FOR u := 1 TO GVL_PARAM.UNIT_COUNT DO
	_stOut.astUnit[u].bPSetActive := FALSE;
END_FOR
IF i_nUnit >= 1 AND i_nUnit <= GVL_PARAM.UNIT_COUNT THEN
	_stOut.astUnit[i_nUnit].bPSetActive	:= i_bUnitPSetActive;
	_stOut.astUnit[i_nUnit].fPSet		:= i_fUnitPSet;
END_IF
// 새 지령: 값이 바뀌었거나 i_bSend
// [결함 13 수정 2026-11-04: 값 비교를 비트로 (운전원이 NaN을 넣어도 여기서 멈추지 않고 고르기에서 이상값으로 거름). 원래 _stOut.fPSet <> stOld.fPSet, _stOut.fQSet <> stOld.fQSet, …fPSet <> stOld.astUnit[u].fPSet]
_stOut.bNewSet := i_bSend
	OR _stOut.bPSetActive <> stOld.bPSetActive OR F_RealChanged(_stOut.fPSet, stOld.fPSet)
	OR _stOut.bQSetActive <> stOld.bQSetActive OR F_RealChanged(_stOut.fQSet, stOld.fQSet);
FOR u := 1 TO GVL_PARAM.UNIT_COUNT DO
	_stOut.bNewSet := _stOut.bNewSet
		OR _stOut.astUnit[u].bPSetActive <> stOld.astUnit[u].bPSetActive
		OR F_RealChanged(_stOut.astUnit[u].fPSet, stOld.astUnit[u].fPSet);
END_FOR
i_bSend := FALSE;

M_UpdateOutput := TRUE;		// 시험용: 항상 살아 있음 (만료 없음)
END_METHOD

END_FUNCTION_BLOCK

// ---- 20_Module/ControlMode/FB_CmPeakCut.TcPOU
FUNCTION_BLOCK FB_CmPeakCut EXTENDS FB_CmTariffBase		// 제어 모드: 피크컷 (Messis PEAK_SHAVING_MODE). 15분 평균 수전이 목표를 넘지 않게 방전
// 우선순위: 자동 충전 시간 → 잔량 방전 시간 (잔량 방전과 피크 제어 중 큰 값, 방전 허용 시간에만) → 피크 제어 (방전 허용 시간에만). 휴일·시각 무효 → 0
// 방전은 모두 역송 방지 (공통 설정). 피크 제어량 계산은 FB_CmPeakCalc (통합 모드와 같음)
VAR_INPUT
	i_stSet		: ST_CmPeakCutSet;		// 설정 (A_PassModuleSet이 GVL_PERSIST.g_stModuleSet.stCmPeakCut을 매 스캔 넘김)
END_VAR
VAR_OUTPUT
	q_fPeakCtrl	: REAL;		// 진단: 피크 제어량 (kW, FB_CmPeakCalc)
	q_nRemainMin	: UINT;		// 진단: 15분 구간 남은 분
	q_fExceeded	: REAL;		// 진단: 구간 목표 초과 수전 누적 (kW·분)
	q_fLoad1m	: REAL;		// 진단: 직전 1분 평균 부하 (kW)
END_VAR
VAR
	_fbPeak		: FB_CmPeakCalc;
END_VAR

METHOD M_Enter
VAR_INPUT
	i_stView	: ST_CtrlModeView;
END_VAR
SUPER^.M_Enter(i_stView := i_stView);
_fbPeak.M_Reset();
END_METHOD

METHOD M_Calc : ST_CtrlModeOut
VAR_INPUT
	i_stView	: ST_CtrlModeView;
END_VAR
VAR
	nNow	: UINT;
	fP		: REAL;
	fRem	: REAL;
	nRsn	: UINT;
	bNoCap	: BOOL;
END_VAR
fP := 0.0;
_fbPeak(i_stSet := i_stSet.stPeak, i_fRevMargin := i_stCommon.stNoRev.fMargin, i_stView := i_stView);		// 휴일에도 평균은 셈
q_fPeakCtrl		:= _fbPeak.q_fCtrl;
q_nRemainMin	:= _fbPeak.q_nRemainMin;
q_fExceeded		:= _fbPeak.q_fExceeded;
q_fLoad1m		:= _fbPeak.q_fLoad1m;
IF M_Begin(i_stView := i_stView) THEN
	nNow := F_TimeHhmm(i_stTime := i_stView.stTime);
	IF i_stSet.stAutoChg.bUse AND F_InHhmmWindow(i_nNow := nNow, i_nStart := i_stSet.stAutoChg.nStart, i_nEnd := i_stSet.stAutoChg.nEnd) THEN
		// 1) 자동 충전 (Messis MT_auto_charge)
		fP			:= -M_AutoChg(i_stView := i_stView, i_stWin := i_stSet.stAutoChg, q_bNoCap => bNoCap);
		q_nState	:= SEL(bNoCap, GVL_CM_RSN.AUTO_CHG, GVL_CM_RSN.NO_CAP);
	ELSIF i_stSet.stRemain.bUse AND F_InHhmmWindow(i_nNow := nNow, i_nStart := i_stSet.stRemain.nStart, i_nEnd := i_stSet.stRemain.nEnd) THEN
		// 2) 잔량 방전 (Messis MT_remain_discharge): 잔량 방전량이 있을 때만, 피크 제어량이 더 크면 그 값
		// [14번 수정 2026-11-09: 방전 허용 시간(공통 stDis: 시간·일요일) 밖이면 잔량 방전·피크 제어 모두 0, 상태 DIS_TIME.
		//   원래는 잔량 방전 시간이면 방전 허용 시간을 보지 않고 방전함]
		IF NOT M_DisAllowed(i_stTime := i_stView.stTime) THEN
			q_nState := GVL_CM_RSN.DIS_TIME;
		ELSE
			fRem		:= M_RemainDis(i_stView := i_stView, i_stWin := i_stSet.stRemain, q_bNoCap => bNoCap);
			q_nState	:= SEL(bNoCap, GVL_CM_RSN.REMAIN_DIS, GVL_CM_RSN.NO_CAP);
			IF fRem > 0.0 THEN
				fP := M_NoReverse(i_fReq := MAX(fRem, _fbPeak.q_fCtrl), i_stView := i_stView, q_nRsn => nRsn);
				IF nRsn <> 0 THEN
					q_nState := nRsn;
				END_IF
			END_IF
		END_IF
	ELSIF _fbPeak.q_bNewInterval THEN
		q_nState := GVL_CM_RSN.NEW_INTERVAL;
	ELSIF _fbPeak.q_fCtrl <= 0.0 THEN
		q_nState := GVL_CM_RSN.BELOW_PEAK;
	ELSIF NOT M_DisAllowed(i_stTime := i_stView.stTime) THEN
		q_nState := GVL_CM_RSN.DIS_TIME;
	ELSE
		// 3) 피크 제어 (Messis MT_peak_shaving_mode)
		fP			:= M_NoReverse(i_fReq := _fbPeak.q_fCtrl, i_stView := i_stView, q_nRsn => nRsn);
		q_nState	:= SEL(nRsn <> 0, GVL_CM_RSN.PEAK, nRsn);
	END_IF
END_IF
M_Calc := M_Finish(i_fP := fP);
END_METHOD

METHOD M_CheckSet : WSTRING(63)
M_CheckSet := SUPER^.M_CheckSet();
IF M_CheckSet <> "" THEN
	RETURN;
END_IF
// [결함 13 수정 2026-11-04: 피크 설정이 숫자인지 먼저]
IF NOT (F_RealOk(i_stSet.stPeak.fTarget) AND F_RealOk(i_stSet.stPeak.fBandSens) AND F_RealOk(i_stSet.stPeak.fLoadRatio) AND F_RealOk(i_stSet.stPeak.fMinOut)) THEN
	M_CheckSet := "피크컷: 피크 설정 숫자 아님";
ELSIF i_stSet.stPeak.fTarget < 0.0 OR i_stSet.stPeak.fBandSens < 0.0 OR i_stSet.stPeak.fLoadRatio < 0.0 OR i_stSet.stPeak.fLoadRatio > 1.0 OR i_stSet.stPeak.fMinOut < 0.0 THEN
	M_CheckSet := "피크컷: 목표·감도·부하 비율(0~1)·최소 출력";
ELSIF NOT M_CheckWindow(i_stWin := i_stSet.stAutoChg) THEN
	M_CheckSet := "피크컷: 자동 충전 시간·SOC";
ELSIF NOT M_CheckWindow(i_stWin := i_stSet.stRemain) THEN
	M_CheckSet := "피크컷: 잔량 방전 시간·SOC";
END_IF
END_METHOD

END_FUNCTION_BLOCK

// ---- 20_Module/ControlMode/FB_CmPeakCalc.TcPOU
FUNCTION_BLOCK FB_CmPeakCalc		// 15분 피크 제어량 계산 (Messis ACT_calc_quarter_avg_and_output 이식). 피크컷·통합 모드가 같이 씀
// 구간 = 시계 기준 15분 (매시 00·15·30·45분). 1초마다 수전·부하 평균, 시계 분이 바뀔 때마다 제어량 갱신, 구간 경계에서 0:
//   목표를 넘은 수전 누적 / 남은 분 (10 단위 반올림) × 속도 × (지난 분/15), 가용 출력 · 30초 평균 부하 × fLoadRatio · (30초 평균 부하 − 역송 여유) 상한
// 켜진 모드에서 매 스캔 부름. 모드가 켜질 때 M_Reset
VAR_INPUT
	i_stSet			: ST_CmPeakCalcSet;
	i_fRevMargin	: REAL;				// kW, 역송 방지 여유 (공통 설정 stNoRev.fMargin)
	i_stView		: ST_CtrlModeView;
END_VAR
VAR_OUTPUT
	q_fCtrl			: REAL;		// kW, 피크 제어 방전량 (0 = 제어 안 함). 1분마다 바뀜
	q_bNewInterval	: BOOL;		// 이번 스캔에 새 15분 구간 시작 (1스캔)
	q_nRemainMin	: UINT;		// 구간 남은 분
	q_fExceeded		: REAL;		// 이 구간 목표를 넘은 수전 누적 (kW·분)
	q_fLoad1m		: REAL;		// 직전 1분 평균 부하 (kW, ESS가 없을 때의 수전)
	q_bNoPcc		: BOOL;		// 접속점 계측 무효 (제어량 0, 평균 안 셈)
END_VAR
VAR
	_bInit			: BOOL;
	_nQuarter		: UINT;		// 지금 구간 번호 (시 × 4 + 분 / 15)
	_nPrevSec		: UINT;		// 지난 스캔 시계 초
	_nPrevMin		: UINT;		// 지난 스캔 시계 분
	_nPrevHalf		: UINT;		// 지난 스캔 30초 칸 (0 / 1)
	_n60			: UINT;		// 1분 평균 표본 수
	_n30			: UINT;		// 30초 평균 표본 수
	_fImp1m			: REAL;		// 1분 평균 수전 (kW)
	_fLoad30		: REAL;		// 30초 평균 부하 (kW)
	_fVelocity		: REAL;		// 제어 속도 (F_CmVelocity)
END_VAR
VAR_TEMP
	nQ				: UINT;
	fImp			: REAL;		// 수전 (kW)
	fLoad			: REAL;		// 부하 (kW)
	fCtrl			: REAL;
	nMin			: UINT;		// 구간 시작부터 지난 분
END_VAR

q_bNewInterval := FALSE;
q_bNoPcc := NOT i_stView.stGroup.stPcc.stMeas.stP.bValid;
IF NOT i_stView.stTime.bValid OR i_stSet.fTarget <= 0.0 THEN
	q_fCtrl	:= 0.0;
	_bInit	:= FALSE;
	RETURN;
END_IF

// 1) 구간 시작 (처음 또는 15분 경계). 경계에서는 제어량 0 (Messis: 남은 분 0으로 계산해 0)
nQ := i_stView.stTime.nHour * 4 + i_stView.stTime.nMinute / 15;
IF NOT _bInit OR nQ <> _nQuarter THEN
	q_bNewInterval	:= _bInit;		// 모드가 켜진 첫 스캔은 새 구간으로 보지 않음
	_bInit			:= TRUE;
	_nQuarter		:= nQ;
	_nPrevSec		:= i_stView.stTime.nSecond;
	_nPrevMin		:= i_stView.stTime.nMinute;
	_nPrevHalf		:= i_stView.stTime.nSecond / 30;
	_n60			:= 0;
	_n30			:= 0;
	q_nRemainMin	:= 15 - i_stView.stTime.nMinute MOD 15;
	q_fExceeded		:= 0.0;
	q_fCtrl			:= 0.0;
	_fVelocity		:= F_CmVelocity(i_fH := i_stSet.fTarget);
	RETURN;
END_IF

// 2) 시계의 초가 바뀔 때마다 (분·30초 경계는 시계 값으로 판단: 시계 보정으로 초가 건너뛰어도 밀리지 않음)
IF i_stView.stTime.nSecond <> _nPrevSec THEN
	_nPrevSec := i_stView.stTime.nSecond;
	// 3) 분이 바뀌면 지난 1분 평균으로 제어량 갱신
	IF i_stView.stTime.nMinute <> _nPrevMin THEN
		_nPrevMin		:= i_stView.stTime.nMinute;
		nMin			:= i_stView.stTime.nMinute MOD 15;		// 구간 시작부터 지난 분
		q_nRemainMin	:= 15 - nMin;
		fCtrl			:= 0.0;
		IF _n60 > 0 AND NOT q_bNoPcc THEN
			q_fExceeded := q_fExceeded + (_fImp1m - i_stSet.fTarget);
			IF q_fLoad1m - i_stSet.fTarget > i_stView.stGroup.fPRatedAvail * UINT_TO_REAL(q_nRemainMin / 15) * i_stSet.fBandSens * 0.5 THEN
				fCtrl := MIN(F_CmRoundTens(i_f := q_fExceeded / UINT_TO_REAL(q_nRemainMin)) * _fVelocity * (UINT_TO_REAL(nMin) / 15.0), i_stView.stGroup.fPRatedAvail);
			END_IF
			fCtrl := MIN(fCtrl, _fLoad30 * i_stSet.fLoadRatio);
			fCtrl := MIN(fCtrl, _fLoad30 - i_fRevMargin);
			IF fCtrl <= 1.0 THEN
				fCtrl := 0.0;
			ELSE
				fCtrl := MAX(fCtrl, i_stSet.fMinOut);
			END_IF
			IF _fImp1m - i_stSet.fTarget > 0.0 THEN
				_fVelocity := F_CmVelocity(i_fH := _fImp1m - i_stSet.fTarget);
			END_IF
		END_IF
		q_fCtrl	:= fCtrl;
		_n60	:= 0;			// 다음 1분 평균을 새로 셈 (값은 남김)
	END_IF
	IF i_stView.stTime.nSecond / 30 <> _nPrevHalf THEN
		_nPrevHalf	:= i_stView.stTime.nSecond / 30;
		_n30		:= 0;		// 다음 30초 평균을 새로 셈 (값은 남김)
	END_IF
	// 4) 1초 표본
	IF q_bNoPcc THEN
		q_fCtrl := 0.0;			// 계측 무효: 평균에 넣지 않고 제어 안 함
	ELSE
		_n60	:= _n60 + 1;
		_n30	:= _n30 + 1;
		fImp	:= -i_stView.stGroup.stPcc.stMeas.stP.fValue;			// 수전 + (접속점 P는 공급 +)
		fLoad	:= i_stView.stGroup.fPOut + fImp;							// ESS가 없을 때의 수전
		_fImp1m		:= (_fImp1m * UINT_TO_REAL(_n60 - 1) + fImp) / UINT_TO_REAL(_n60);
		q_fLoad1m	:= (q_fLoad1m * UINT_TO_REAL(_n60 - 1) + fLoad) / UINT_TO_REAL(_n60);
		_fLoad30	:= (_fLoad30 * UINT_TO_REAL(_n30 - 1) + fLoad) / UINT_TO_REAL(_n30);
	END_IF
END_IF

METHOD M_Reset		// 모드가 켜질 때: 구간을 지금부터 다시 셈, 제어량 0
_bInit		:= FALSE;
q_fCtrl		:= 0.0;
q_fExceeded	:= 0.0;
q_fLoad1m	:= 0.0;
_fImp1m		:= 0.0;
_fLoad30	:= 0.0;
END_METHOD

END_FUNCTION_BLOCK

// ---- 20_Module/ControlMode/F_CmVelocity.TcPOU
FUNCTION F_CmVelocity : REAL		// 피크 제어 속도 (Messis getVelocity): 넘는 양이 작을수록 크게. (log10(h + 100) − log10(h)) × 20, h ≤ 0이면 1
VAR_INPUT
	i_fH		: REAL;		// kW, 목표 또는 목표를 넘은 양
END_VAR

IF i_fH <= 0.0 THEN
	F_CmVelocity := 1.0;
ELSE
	F_CmVelocity := (LOG(i_fH + 100.0) - LOG(i_fH)) * 20.0;
END_IF

END_FUNCTION

// ---- 20_Module/ControlMode/F_CmRoundTens.TcPOU
FUNCTION F_CmRoundTens : REAL		// 10 단위 반올림 (Messis roundUpTens)
VAR_INPUT
	i_f			: REAL;
END_VAR

// [결함 13 수정 2026-11-04: NaN·범위 밖이면 REAL_TO_DINT가 FPU 예외 → F_RealToDint (NaN은 0). 원래 DINT_TO_REAL(REAL_TO_DINT(i_f / 10.0)) * 10.0]
F_CmRoundTens := DINT_TO_REAL(F_RealToDint(i_f / 10.0)) * 10.0;

END_FUNCTION

// ---- 20_Module/ControlMode/FB_CmSchedPeak.TcPOU
FUNCTION_BLOCK FB_CmSchedPeak EXTENDS FB_CmTariffBase		// 제어 모드: 통합 = 스케줄 + 피크컷 (Messis SCHEDULE_PS_MODE)
// 우선순위: 잔량 방전 시간 (잔량 방전과 피크 제어 중 큰 값, 방전 허용 시간에만) → 피크 제어가 필요하고 방전 허용 시간이면 (피크 제어량과 시간표 방전 중 큰 값)
//   → 아니면 스케줄 모드와 같음. 시간표는 스케줄 모드와 같은 표, 피크 제어량 계산은 피크컷과 같은 FB_CmPeakCalc
// Messis와 다른 점: 시간표가 충전 칸일 때 피크 제어가 필요하면 피크 제어량만 방전 (Messis는 충전값 크기만큼 방전할 수 있었음)
VAR_INPUT
	i_stTable	: ST_CmScheduleSet;		// 시간표 (스케줄 모드와 같은 GVL_PERSIST.g_stModuleSet.stCmSchedule)
	i_stSet		: ST_CmSchedPeakSet;	// 설정 (GVL_PERSIST.g_stModuleSet.stCmSchedPeak)
END_VAR
VAR_OUTPUT
	q_fPeakCtrl	: REAL;		// 진단: 피크 제어량 (kW, FB_CmPeakCalc)
	q_nRemainMin	: UINT;		// 진단: 15분 구간 남은 분
	q_fExceeded	: REAL;		// 진단: 구간 목표 초과 수전 누적 (kW·분)
	q_fLoad1m	: REAL;		// 진단: 직전 1분 평균 부하 (kW)
END_VAR
VAR
	_fbPeak		: FB_CmPeakCalc;
END_VAR

METHOD M_Enter
VAR_INPUT
	i_stView	: ST_CtrlModeView;
END_VAR
SUPER^.M_Enter(i_stView := i_stView);
_fbPeak.M_Reset();
END_METHOD

METHOD M_Calc : ST_CtrlModeOut
VAR_INPUT
	i_stView	: ST_CtrlModeView;
END_VAR
VAR
	nNow	: UINT;
	fP		: REAL;
	fRem	: REAL;
	nRsn	: UINT;
	bNoCap	: BOOL;
END_VAR
fP := 0.0;
_fbPeak(i_stSet := i_stSet.stPeak, i_fRevMargin := i_stCommon.stNoRev.fMargin, i_stView := i_stView);
q_fPeakCtrl		:= _fbPeak.q_fCtrl;
q_nRemainMin	:= _fbPeak.q_nRemainMin;
q_fExceeded		:= _fbPeak.q_fExceeded;
q_fLoad1m		:= _fbPeak.q_fLoad1m;
IF M_Begin(i_stView := i_stView) THEN
	nNow := F_TimeHhmm(i_stTime := i_stView.stTime);
	M_SchedLookup(i_stTime := i_stView.stTime, iq_stTable := i_stTable);
	IF i_stSet.stRemain.bUse AND F_InHhmmWindow(i_nNow := nNow, i_nStart := i_stSet.stRemain.nStart, i_nEnd := i_stSet.stRemain.nEnd) THEN
		// 1) 잔량 방전
		// [14번 수정 2026-11-09: 방전 허용 시간(공통 stDis: 시간·일요일) 밖이면 잔량 방전·피크 제어 모두 0, 상태 DIS_TIME.
		//   원래는 잔량 방전 시간이면 방전 허용 시간을 보지 않고 방전함]
		IF NOT M_DisAllowed(i_stTime := i_stView.stTime) THEN
			q_nState := GVL_CM_RSN.DIS_TIME;
		ELSE
			fRem		:= M_RemainDis(i_stView := i_stView, i_stWin := i_stSet.stRemain, q_bNoCap => bNoCap);
			q_nState	:= SEL(bNoCap, GVL_CM_RSN.REMAIN_DIS, GVL_CM_RSN.NO_CAP);
			IF fRem > 0.0 THEN
				fP := M_NoReverse(i_fReq := MAX(fRem, _fbPeak.q_fCtrl), i_stView := i_stView, q_nRsn => nRsn);
				IF nRsn <> 0 THEN
					q_nState := nRsn;
				END_IF
			END_IF
		END_IF
	ELSIF _fbPeak.q_fCtrl > 0.0 AND M_DisAllowed(i_stTime := i_stView.stTime) THEN
		// 2) 피크 제어 + 시간표 방전 중 큰 값
		fP			:= M_NoReverse(i_fReq := MAX(_fbPeak.q_fCtrl, MAX(q_fSlotP, 0.0)), i_stView := i_stView, q_nRsn => nRsn);
		q_nState	:= SEL(nRsn <> 0, GVL_CM_RSN.SCHED_PEAK, nRsn);
	ELSE
		// 3) 스케줄만
		fP			:= M_SchedOut(i_stView := i_stView, q_nRsn => nRsn);
		q_nState	:= nRsn;
	END_IF
END_IF
M_Calc := M_Finish(i_fP := fP);
END_METHOD

METHOD M_CheckSet : WSTRING(63)
M_CheckSet := SUPER^.M_CheckSet();
IF M_CheckSet <> "" THEN
	RETURN;
END_IF
M_CheckSet := M_CheckTable(iq_stTable := i_stTable);
IF M_CheckSet <> "" THEN
	RETURN;
END_IF
// [결함 13 수정 2026-11-04: 피크 설정이 숫자인지 먼저]
IF NOT (F_RealOk(i_stSet.stPeak.fTarget) AND F_RealOk(i_stSet.stPeak.fBandSens) AND F_RealOk(i_stSet.stPeak.fLoadRatio) AND F_RealOk(i_stSet.stPeak.fMinOut)) THEN
	M_CheckSet := "통합: 피크 설정 숫자 아님";
ELSIF i_stSet.stPeak.fTarget < 0.0 OR i_stSet.stPeak.fBandSens < 0.0 OR i_stSet.stPeak.fLoadRatio < 0.0 OR i_stSet.stPeak.fLoadRatio > 1.0 OR i_stSet.stPeak.fMinOut < 0.0 THEN
	M_CheckSet := "통합: 목표·감도·부하 비율(0~1)·최소 출력";
ELSIF NOT M_CheckWindow(i_stWin := i_stSet.stRemain) THEN
	M_CheckSet := "통합: 잔량 방전 시간·SOC";
END_IF
END_METHOD

END_FUNCTION_BLOCK

// ---- 20_Module/Common/FB_SocLimit.TcPOU
FUNCTION_BLOCK FB_SocLimit EXTENDS FB_ModuleBase IMPLEMENTS I_BatLimitRule	// SOC 감발·차단·재개 마진 (버스 제한). 기본 SOC 정책 (Auto·Manual 기본 등록)
// 최대 SOC가 상한에 다가가면 충전 한도를, 최소 SOC가 하한에 다가가면 방전 한도를 줄이고, 한계에서 막음
// 막은 뒤에는 SOC가 재개 마진만큼 돌아와야 다시 허용. 다시 허용한 뒤 감발 구간을 지나는 동안 bResume (재개 램프율)
// 출력 한도만 냄 (장비 명령 없음). 한도가 0이면 그 방향 출력 0 = 대기
// nTarget 0 = 모든 버스를 한 인스턴스가 봄 (버스마다 상태를 따로 가짐)
VAR_INPUT
	i_stSet	: ST_SocLimitSet;	// 설정 (MAIN이 GVL_PERSIST.g_stModuleSet 칸을 매 스캔 넘김. 안 넘기면 기본값)
END_VAR
VAR
	(* 버스마다 상태 *)
	_abChgBlock	: ARRAY[1..GVL_PARAM.BAT_COUNT] OF BOOL;	// 충전 막음 (재개 마진 전까지 유지)
	_abDisBlock	: ARRAY[1..GVL_PARAM.BAT_COUNT] OF BOOL;	// 방전 막음
	_abChgResume	: ARRAY[1..GVL_PARAM.BAT_COUNT] OF BOOL;	// 충전 재개 중 (막음이 풀린 뒤 감발 구간)
	_abDisResume	: ARRAY[1..GVL_PARAM.BAT_COUNT] OF BOOL;
	_afChgRatio	: ARRAY[1..GVL_PARAM.BAT_COUNT] OF REAL;	// 진단: 충전 한도 비율 (1 = 안 줄임)
	_afDisRatio	: ARRAY[1..GVL_PARAM.BAT_COUNT] OF REAL;	// 진단: 방전 한도 비율
END_VAR
VAR CONSTANT
	RSN_CHG_DERATE	: UINT := 1;	// 상한 근처 충전 감발
	RSN_CHG_BLOCK	: UINT := 2;	// 상한 충전 막음
	RSN_DIS_DERATE	: UINT := 3;	// 하한 근처 방전 감발
	RSN_DIS_BLOCK	: UINT := 4;	// 하한 방전 막음
	RSN_SOC_INVALID	: UINT := 5;	// SOC 무효
END_VAR

METHOD M_Evaluate : ST_BatLimitOut
VAR_INPUT
	i_stView	: ST_BatLimitView;
END_VAR
VAR
	b	: UINT;
	fChg	: REAL;	// 충전 한도 비율
	fDis	: REAL;	// 방전 한도 비율
END_VAR
b := i_stView.nBatGroup;
IF b < 1 OR b > GVL_PARAM.BAT_COUNT THEN
	RETURN;
END_IF
// SOC 무효: 상태를 풀고, 설정이면 충·방전 모두 막음
IF NOT i_stView.stSocMax.bValid OR NOT i_stView.stSocMin.bValid THEN
	_abChgBlock[b]	:= FALSE;
	_abDisBlock[b]	:= FALSE;
	_abChgResume[b]	:= FALSE;
	_abDisResume[b]	:= FALSE;
	_afChgRatio[b]	:= 1.0;
	_afDisRatio[b]	:= 1.0;
	IF i_stSet.bBlockOnInvalid THEN
		M_Evaluate.stP.bActive	:= TRUE;
		M_Evaluate.stP.fMax	:= 0.0;
		M_Evaluate.stP.fMin	:= 0.0;
		M_Evaluate.stP.nReason	:= RSN_SOC_INVALID;
		_afChgRatio[b]	:= 0.0;
		_afDisRatio[b]	:= 0.0;
	END_IF
	RETURN;
END_IF

// 충전: 최대 SOC 기준
IF i_stView.stSocMax.fValue >= i_stSet.fSocMax THEN
	_abChgBlock[b]	:= TRUE;
	_abChgResume[b]	:= FALSE;
ELSIF _abChgBlock[b] AND i_stView.stSocMax.fValue <= i_stSet.fSocMax - i_stSet.fResumeMargin THEN
	_abChgBlock[b]	:= FALSE;
	_abChgResume[b]	:= TRUE;
END_IF
fChg := 0.0;
IF NOT _abChgBlock[b] THEN
	fChg := F_SocDerate(i_fSoc := i_stView.stSocMax.fValue, i_fLimit := i_stSet.fSocMax, i_fBand := i_stSet.fBand, i_bUpper := TRUE);
END_IF
IF fChg >= 1.0 THEN
	_abChgResume[b] := FALSE;
END_IF

// 방전: 최소 SOC 기준
IF i_stView.stSocMin.fValue <= i_stSet.fSocMin THEN
	_abDisBlock[b]	:= TRUE;
	_abDisResume[b]	:= FALSE;
ELSIF _abDisBlock[b] AND i_stView.stSocMin.fValue >= i_stSet.fSocMin + i_stSet.fResumeMargin THEN
	_abDisBlock[b]	:= FALSE;
	_abDisResume[b]	:= TRUE;
END_IF
fDis := 0.0;
IF NOT _abDisBlock[b] THEN
	fDis := F_SocDerate(i_fSoc := i_stView.stSocMin.fValue, i_fLimit := i_stSet.fSocMin, i_fBand := i_stSet.fBand, i_bUpper := FALSE);
END_IF
IF fDis >= 1.0 THEN
	_abDisResume[b] := FALSE;
END_IF

_afChgRatio[b]	:= fChg;
_afDisRatio[b]	:= fDis;
M_Evaluate.bResume := _abChgResume[b] OR _abDisResume[b];
IF fChg < 1.0 OR fDis < 1.0 THEN
	M_Evaluate.stP.bActive	:= TRUE;
	M_Evaluate.stP.fMax	:= MAX(i_stView.fPDisMax, 0.0) * fDis;
	M_Evaluate.stP.fMin	:= -MAX(i_stView.fPChgMax, 0.0) * fChg;
	// 이유: 막음이 감발보다 먼저 (한 줄 제한이라 상·하한이 같은 이유를 가짐)
	IF _abDisBlock[b] THEN
		M_Evaluate.stP.nReason := RSN_DIS_BLOCK;
	ELSIF _abChgBlock[b] THEN
		M_Evaluate.stP.nReason := RSN_CHG_BLOCK;
	ELSIF fDis < 1.0 THEN
		M_Evaluate.stP.nReason := RSN_DIS_DERATE;
	ELSE
		M_Evaluate.stP.nReason := RSN_CHG_DERATE;
	END_IF
END_IF
END_METHOD

METHOD M_ReasonText : WSTRING(63)
VAR_INPUT
	i_nReason	: UINT;
END_VAR
CASE i_nReason OF
	RSN_CHG_DERATE:	M_ReasonText := "SOC 상한 근처 충전 감발";
	RSN_CHG_BLOCK:	M_ReasonText := "SOC 상한 충전 막음";
	RSN_DIS_DERATE:	M_ReasonText := "SOC 하한 근처 방전 감발";
	RSN_DIS_BLOCK:	M_ReasonText := "SOC 하한 방전 막음";
	RSN_SOC_INVALID:	M_ReasonText := "SOC 무효";
ELSE
	M_ReasonText := WCONCAT("이유 ", TO_WSTRING(i_nReason));
END_CASE
END_METHOD

METHOD M_CheckSet : WSTRING(63)		// 설정 점검: SOC 상·하한, 감발 폭, 재개 마진
// [9-21 수정 2026-11-04: 검사 규칙을 F_SocLimitSetErr로 옮김 (EMS config 반영 FB_EmsConfigApply와 같은 규칙을 씀). 원래:
//   M_CheckSet := "";
//   IF NOT (F_RealOk(i_stSet.fSocMin) AND F_RealOk(i_stSet.fSocMax) AND F_RealOk(i_stSet.fBand) AND F_RealOk(i_stSet.fResumeMargin)) THEN	// [결함 13 수정 2026-11-04]
//   	M_CheckSet := "SOC 설정 숫자 아님";
//   ELSIF i_stSet.fSocMin < 0.0 OR i_stSet.fSocMax > 100.0 OR i_stSet.fSocMin >= i_stSet.fSocMax THEN
//   	M_CheckSet := "SOC 상·하한 (0 ≤ 하한 < 상한 ≤ 100)";
//   ELSIF i_stSet.fBand < 0.0 OR i_stSet.fSocMin + i_stSet.fBand > i_stSet.fSocMax - i_stSet.fBand THEN
//   	M_CheckSet := "감발 폭 fBand (0 이상, 상·하한 사이)";
//   ELSIF i_stSet.fResumeMargin < 0.0 OR i_stSet.fSocMin + i_stSet.fResumeMargin >= i_stSet.fSocMax - i_stSet.fResumeMargin THEN
//   	M_CheckSet := "재개 마진 fResumeMargin (0 이상, 상·하한 사이)";
//   END_IF]
M_CheckSet := F_SocLimitSetErr(i_stSet);
END_METHOD

END_FUNCTION_BLOCK

// ---- 20_Module/Common/F_SocDerate.TcPOU
FUNCTION F_SocDerate : REAL	// SOC 감발 비율 (0~1, 상태 없음). 여러 SOC 정책 모듈이 같이 씀
// 상한(i_bUpper = TRUE, 충전 쪽): SOC ≥ 한계면 0, 한계 - 폭 < SOC면 선형으로 줄임, 그 아래는 1
// 하한(i_bUpper = FALSE, 방전 쪽): SOC ≤ 한계면 0, SOC < 한계 + 폭이면 선형으로 줄임, 그 위는 1
VAR_INPUT
	i_fSoc	: REAL;	// %
	i_fLimit	: REAL;	// %, 한계
	i_fBand	: REAL;	// %, 감발 폭. 0 이하면 줄이지 않고 한계에서 0
	i_bUpper	: BOOL;	// TRUE = 상한, FALSE = 하한
END_VAR

IF i_bUpper THEN
	IF i_fSoc >= i_fLimit THEN
		F_SocDerate := 0.0;
	ELSIF i_fBand > 0 AND i_fSoc > i_fLimit - i_fBand THEN
		F_SocDerate := (i_fLimit - i_fSoc) / i_fBand;
	ELSE
		F_SocDerate := 1.0;
	END_IF
ELSE
	IF i_fSoc <= i_fLimit THEN
		F_SocDerate := 0.0;
	ELSIF i_fBand > 0 AND i_fSoc < i_fLimit + i_fBand THEN
		F_SocDerate := (i_fSoc - i_fLimit) / i_fBand;
	ELSE
		F_SocDerate := 1.0;
	END_IF
END_IF

END_FUNCTION

// ---- 20_Module/Common/FB_UnitLimit.TcPOU
FUNCTION_BLOCK FB_UnitLimit EXTENDS FB_ModuleBase IMPLEMENTS I_UnitLimitRule	// 사용자 한도: 유닛마다 운전원이 정한 P·Q 상·하한 (kW·kvar). 정격·Derate와 겹쳐 좁은 쪽 (코어 FB_EquipmentLimits)
// 등록: g_aipUnitRule 한 칸, g_astUnitRuleReg nTarget 0 (전체 유닛, 유닛마다 설정을 따로 봄), bAuto·bManual로 적용 모드
// 출력 제한 이유: 유닛 한도 UnitRule + 이 모듈 ID, 이유 "사용자 한도"
VAR_INPUT
	i_stSet		: ST_UnitLimitSet;	// 유닛마다 한도 (MAIN A_PassModuleSet이 g_stModuleSet 칸을 넘김. 안 넘기면 모두 끔)
END_VAR
VAR CONSTANT
	RSN_USER	: UINT := 1;		// 사용자 한도
END_VAR

METHOD M_Evaluate : ST_LimitOut
VAR_INPUT
	i_stView	: ST_UnitLimitView;
END_VAR
VAR
	u	: UINT;
END_VAR
u := i_stView.nUnit;
IF u < 1 OR u > GVL_PARAM.UNIT_COUNT THEN
	RETURN;
END_IF
IF i_stSet.astUnit[u].bPEnable THEN
	M_Evaluate.stP.bActive	:= TRUE;
	M_Evaluate.stP.fMax		:= i_stSet.astUnit[u].fPMax;
	M_Evaluate.stP.fMin		:= i_stSet.astUnit[u].fPMin;
	M_Evaluate.stP.nReason	:= RSN_USER;
END_IF
IF i_stSet.astUnit[u].bQEnable THEN
	M_Evaluate.stQ.bActive	:= TRUE;
	M_Evaluate.stQ.fMax		:= i_stSet.astUnit[u].fQMax;
	M_Evaluate.stQ.fMin		:= i_stSet.astUnit[u].fQMin;
	M_Evaluate.stQ.nReason	:= RSN_USER;
END_IF
END_METHOD

METHOD M_ReasonText : WSTRING(63)
VAR_INPUT
	i_nReason	: UINT;
END_VAR
IF i_nReason = RSN_USER THEN
	M_ReasonText := "사용자 한도";
ELSE
	M_ReasonText := WCONCAT("이유 ", TO_WSTRING(i_nReason));
END_IF
END_METHOD

METHOD M_CheckSet : WSTRING(63)		// 설정 점검: 켠 한도는 상한 ≥ 0 ≥ 하한
VAR
	u	: UINT;
END_VAR
M_CheckSet := "";
FOR u := 1 TO GVL_PARAM.UNIT_COUNT DO
	IF NOT (F_RealOk(i_stSet.astUnit[u].fPMax) AND F_RealOk(i_stSet.astUnit[u].fPMin) AND F_RealOk(i_stSet.astUnit[u].fQMax) AND F_RealOk(i_stSet.astUnit[u].fQMin)) THEN	// [결함 13 수정 2026-11-04]
		M_CheckSet := F_TxtNum("한도 숫자 아님: 유닛 ", u);
		RETURN;
	END_IF
	IF i_stSet.astUnit[u].bPEnable AND (i_stSet.astUnit[u].fPMax < 0.0 OR i_stSet.astUnit[u].fPMin > 0.0) THEN
		M_CheckSet := F_TxtNum("P 한도 상한 < 0 또는 하한 > 0: 유닛 ", u);
		RETURN;
	END_IF
	IF i_stSet.astUnit[u].bQEnable AND (i_stSet.astUnit[u].fQMax < 0.0 OR i_stSet.astUnit[u].fQMin > 0.0) THEN
		M_CheckSet := F_TxtNum("Q 한도 상한 < 0 또는 하한 > 0: 유닛 ", u);
		RETURN;
	END_IF
END_FOR
END_METHOD

END_FUNCTION_BLOCK

// ---- 20_Module/Standard/FB_ProtPcsFault.TcPOU
FUNCTION_BLOCK FB_ProtPcsFault EXTENDS FB_ModuleBase IMPLEMENTS I_ProtectionRule		// 표준 보호: PCS 고장 (범위 Unit): 통신이 있고 PCS가 고장을 알림. 기본 등록. 빼면 이 보호 없음. 현장마다 다르면 복사해 이름을 바꿔 그 칸에 대신 등록
VAR
END_VAR

METHOD M_Evaluate : BOOL		// 범위가 맞지 않게 등록되면 FALSE (보호 안 걸림)
VAR_INPUT
	i_stView	: ST_ProtView;
END_VAR
M_Evaluate := i_stView.eScope = E_ProtScope.Unit AND i_stView.bInstalled AND i_stView.stUnit.bComm AND i_stView.stUnit.bFault;
END_METHOD

END_FUNCTION_BLOCK

// ---- 20_Module/Standard/FB_ProtPcsComm.TcPOU
FUNCTION_BLOCK FB_ProtPcsComm EXTENDS FB_ModuleBase IMPLEMENTS I_ProtectionRule		// 표준 보호: PCS 통신 끊김 (범위 Unit). 기본 등록. 빼면 이 보호 없음. 현장마다 다르면 복사해 이름을 바꿔 그 칸에 대신 등록
VAR
END_VAR

METHOD M_Evaluate : BOOL		// 범위가 맞지 않게 등록되면 FALSE (보호 안 걸림)
VAR_INPUT
	i_stView	: ST_ProtView;
END_VAR
M_Evaluate := i_stView.eScope = E_ProtScope.Unit AND i_stView.bInstalled AND NOT i_stView.stUnit.bComm;
END_METHOD

END_FUNCTION_BLOCK

// ---- 20_Module/Standard/FB_ProtBmsFault.TcPOU
FUNCTION_BLOCK FB_ProtBmsFault EXTENDS FB_ModuleBase IMPLEMENTS I_ProtectionRule		// 표준 보호: BMS 고장 (범위 Bms): 통신이 있고 BMS가 고장을 알림. 기본 등록. 빼면 이 보호 없음. 현장마다 다르면 복사해 이름을 바꿔 그 칸에 대신 등록
VAR
END_VAR

METHOD M_Evaluate : BOOL		// 범위가 맞지 않게 등록되면 FALSE (보호 안 걸림)
VAR_INPUT
	i_stView	: ST_ProtView;
END_VAR
M_Evaluate := i_stView.eScope = E_ProtScope.Bms AND i_stView.bInstalled AND i_stView.stBms.bComm AND i_stView.stBms.bFault;
END_METHOD

END_FUNCTION_BLOCK

// ---- 20_Module/Standard/FB_ProtBmsComm.TcPOU
FUNCTION_BLOCK FB_ProtBmsComm EXTENDS FB_ModuleBase IMPLEMENTS I_ProtectionRule		// 표준 보호: BMS 통신 끊김 (범위 Bms). 기본 등록. 빼면 이 보호 없음. 현장마다 다르면 복사해 이름을 바꿔 그 칸에 대신 등록
VAR
END_VAR

METHOD M_Evaluate : BOOL		// 범위가 맞지 않게 등록되면 FALSE (보호 안 걸림)
VAR_INPUT
	i_stView	: ST_ProtView;
END_VAR
M_Evaluate := i_stView.eScope = E_ProtScope.Bms AND i_stView.bInstalled AND NOT i_stView.stBms.bComm;
END_METHOD

END_FUNCTION_BLOCK

// ---- 20_Module/Standard/FB_ProtPccInvalid.TcPOU
FUNCTION_BLOCK FB_ProtPccInvalid EXTENDS FB_ModuleBase IMPLEMENTS I_ProtectionRule		// 표준 보호: 접속점 계측 무효 (범위 Group): 접속점 유효전력 값이 무효. 기본 등록. 빼면 이 보호 없음. 현장마다 다르면 복사해 이름을 바꿔 그 칸에 대신 등록
VAR
END_VAR

METHOD M_Evaluate : BOOL		// 범위가 맞지 않게 등록되면 FALSE (보호 안 걸림)
VAR_INPUT
	i_stView	: ST_ProtView;
END_VAR
// [결함 7 수정 2026-11-03: 접속점이 없는 그룹(nPccPoint 0)은 판단 안 함. 원래 M_Evaluate := i_stView.eScope = E_ProtScope.Group AND NOT i_stView.stPcc.stMeas.stP.bValid;]
M_Evaluate := i_stView.eScope = E_ProtScope.Group AND NOT i_stView.stPcc.bNoPoint AND NOT i_stView.stPcc.stMeas.stP.bValid;
END_METHOD

END_FUNCTION_BLOCK

// ---- 20_Module/Standard/FB_ProtRespStd.TcPOU
FUNCTION_BLOCK FB_ProtRespStd EXTENDS FB_ModuleBase IMPLEMENTS I_ProtResponse		// 표준 보호 대응 (기본 등록: GVL_SITE.g_aipResp 칸마다 같은 인스턴스): 칸 설정(ST_ProtCfg)의 조치를 범위 안 유닛·BMS에 한 단계로 요청
// 유닛: 범위에 드는 유닛 중 그 운전 모드에 조치를 거는 것(bAuto·bManual)만. 모드 조치(ToManual)는 bAuto 항목이면 범위 안 유닛 전부
// BMS: Bms·BatGroup 범위는 그 버스에 조치를 받는 유닛이 있을 때 (버스에 유닛이 없으면 그대로). Unit·Group·Site 범위는 조치를 받는 유닛의 배터리 그룹 BMS 전부
// 현장 대응이 다르면 이 FB를 복사해 이름을 바꿔 그 칸에 대신 등록. 상태가 없어 인스턴스 하나를 모든 칸에 같이 등록함

METHOD M_Respond		// 칸 설정(stProt)의 조치를 걸렸을 때만 요청
// 코어가 매 스캔 범위 안 대상마다 부름 (조건이 없을 때도: 단계 대응의 타이머·상태를 풀 수 있게). 대상 번호가 0으로 등록되면 대상마다 상태를 따로 둠
VAR_INPUT
	i_bActive		: BOOL;			// 보호 조건 있음 (등록 bAuto·bManual 중 하나가 켜져 있고 조건 모듈이 TRUE)
	i_tActive		: TIME;			// 조건이 이어진 시간 (조건 없으면 0)
	i_nTarget		: UINT;			// 대상 번호 (범위는 i_stRule.eScope. Site면 1)
	i_stRule		: ST_RuleCfg;		// 이 칸 설정 (범위·대상·임계값·표준 대응 설정)
END_VAR
VAR_IN_OUT CONSTANT
	iq_astUnit		: ARRAY[1..GVL_PARAM.UNIT_COUNT] OF ST_UnitState;	// 장비 상태 (이번 스캔 스냅샷, 읽기 전용)
	iq_astBms		: ARRAY[1..GVL_PARAM.BMS_COUNT] OF ST_BatState;
	iq_astUnitCfg	: ARRAY[1..GVL_PARAM.UNIT_COUNT] OF ST_UnitCfg;		// 소속 (제어 그룹·배터리 그룹)
	iq_astBmsCfg	: ARRAY[1..GVL_PARAM.BMS_COUNT] OF ST_BmsCfg;
	iq_aeOpMode		: ARRAY[1..GVL_PARAM.UNIT_COUNT] OF E_OpMode;		// 실제 운전 모드
END_VAR
VAR_IN_OUT
	iq_stReq		: ST_ProtReq;		// 요청 (코어가 비워서 넘김)
END_VAR
VAR
	u			: UINT;
	m			: UINT;
	nBus		: UINT;		// Bms·BatGroup 범위의 배터리 그룹
	nBusUnits	: UINT;		// 그 버스의 유닛 수
	bBusTakes	: BOOL;		// 그 버스에 조치를 받는 유닛이 있음
	bIn			: BOOL;
	bManual		: BOOL;
	bTakes		: BOOL;
	stCfg		: ST_ProtCfg;
END_VAR
IF NOT i_bActive THEN
	RETURN;
END_IF
stCfg := i_stRule.stProt;
nBus := 0;
IF i_stRule.eScope = E_ProtScope.Bms AND i_nTarget >= 1 AND i_nTarget <= GVL_PARAM.BMS_COUNT THEN
	nBus := iq_astBmsCfg[i_nTarget].nBatGroup;
ELSIF i_stRule.eScope = E_ProtScope.BatGroup THEN
	nBus := i_nTarget;
END_IF
(* 1) 유닛 *)
nBusUnits := 0;
bBusTakes := FALSE;
FOR u := 1 TO GVL_PARAM.UNIT_COUNT DO
	CASE i_stRule.eScope OF
		E_ProtScope.Unit:					bIn := u = i_nTarget;
		E_ProtScope.Bms, E_ProtScope.BatGroup:	bIn := nBus <> 0 AND iq_astUnitCfg[u].nBatGroup = nBus;
		E_ProtScope.Group:					bIn := iq_astUnitCfg[u].nGroup = i_nTarget;
		E_ProtScope.Site:					bIn := TRUE;
	ELSE
		bIn := FALSE;
	END_CASE
	IF bIn THEN
		bManual	:= iq_aeOpMode[u] = E_OpMode.Manual;
		bTakes	:= F_ModeApplies(stCfg.bAuto, stCfg.bManual, BOOL_TO_UINT(NOT bManual), BOOL_TO_UINT(bManual));
		nBusUnits := nBusUnits + 1;
		bBusTakes := bBusTakes OR bTakes;
		// 모드 조치: Auto 유닛에 거는 항목이면 실제 모드와 관계없이 (이미 Manual이어도 Auto 재요청을 막음)
		IF stCfg.bAuto AND stCfg.eModeAction = E_ModeAction.ToManual THEN
			iq_stReq.abToManual[u] := TRUE;
		END_IF
		IF bTakes THEN
			iq_stReq.aePcs[u]	:= stCfg.ePcsAction;
			iq_stReq.afPPct[u]	:= stCfg.fPPct;
			iq_stReq.afQPct[u]	:= stCfg.fQPct;
			// 유닛·제어 그룹·사이트 범위: 그 유닛 배터리 그룹의 BMS 전부
			IF stCfg.eBatAction <> E_BatAction.None AND nBus = 0 AND iq_astUnitCfg[u].nBatGroup <> 0 THEN
				FOR m := 1 TO GVL_PARAM.BMS_COUNT DO
					IF iq_astBmsCfg[m].nBatGroup = iq_astUnitCfg[u].nBatGroup THEN
						iq_stReq.aeBat[m] := stCfg.eBatAction;
					END_IF
				END_FOR
			END_IF
		END_IF
	END_IF
END_FOR
(* 2) Bms·BatGroup 범위의 배터리 조치: 버스에 조치를 받는 유닛이 있을 때 (버스에 유닛이 없으면 그대로) *)
IF nBus <> 0 AND stCfg.eBatAction <> E_BatAction.None AND (bBusTakes OR nBusUnits = 0) THEN
	FOR m := 1 TO GVL_PARAM.BMS_COUNT DO
		IF (i_stRule.eScope = E_ProtScope.Bms AND m = i_nTarget) OR (i_stRule.eScope = E_ProtScope.BatGroup AND iq_astBmsCfg[m].nBatGroup = nBus) THEN
			iq_stReq.aeBat[m] := stCfg.eBatAction;
		END_IF
	END_FOR
END_IF
END_METHOD

END_FUNCTION_BLOCK

// ---- 20_Module/Common/FB_RuleValue.TcPOU
FUNCTION_BLOCK FB_RuleValue EXTENDS FB_ModuleBase IMPLEMENTS I_ProtectionRule, I_OutputRule		// 아날로그 값 하나 ↔ 임계값 (온도·습도 등). 임계값은 등록 설정(fThreshold)에서 받음
VAR_INPUT
	i_ipAux			: I_AuxDevice;		// 읽을 보조 장비 (선언 때 지정)
	i_nPoint		: UINT;				// 아날로그 입력 점 번호
	i_stSet			: ST_RuleValueSet;	// 설정: 이하·이상, 해소 폭, 통신 끊김 시 조건 (MAIN이 GVL_PERSIST.g_stModuleSet 칸을 매 스캔 넘김. 안 넘기면 기본값)
END_VAR
VAR
	_bProtCond		: BOOL;				// 보호 규칙 판단 상태 (히스테리시스)
	_bOutCond		: BOOL;				// 출력 규칙 판단 상태 (히스테리시스)
END_VAR

METHOD M_Evaluate : BOOL		// 보호 규칙으로 판단 (보호용 상태 _bProtCond. 값 하나라 대상과 관계없음)
VAR_INPUT
	i_stView	: ST_ProtView;
END_VAR
M_Evaluate := M_Judge(i_fThreshold := i_stView.fThreshold, iq_bCond := _bProtCond);
END_METHOD

METHOD M_Check : BOOL		// 출력 규칙으로 판단 (출력용 상태 _bOutCond. 보호와 같은 인스턴스여도 히스테리시스가 섞이지 않음)
VAR_INPUT
	i_fThreshold	: REAL;
END_VAR
M_Check := M_Judge(i_fThreshold := i_fThreshold, iq_bCond := _bOutCond);
END_METHOD

METHOD PRIVATE M_Judge : BOOL		// 임계값·히스테리시스 판단. 상태는 부르는 쪽 것을 씀
VAR_INPUT
	i_fThreshold	: REAL;
END_VAR
VAR_IN_OUT
	iq_bCond		: BOOL;			// 이 판단의 히스테리시스 상태 (보호용·출력용 따로)
END_VAR
VAR
	stValue			: ST_Val;
END_VAR
IF i_ipAux = 0 THEN
	iq_bCond := FALSE;
ELSE
	stValue := i_ipAux.M_GetValue(i_nPoint);
	IF NOT i_ipAux.Comm OR NOT stValue.bValid THEN
		iq_bCond := i_stSet.bOnCommLoss;
	ELSIF NOT i_stSet.bBelow THEN
		IF stValue.fValue >= i_fThreshold THEN
			iq_bCond := TRUE;
		ELSIF stValue.fValue < i_fThreshold - i_stSet.fHyst THEN
			iq_bCond := FALSE;
		END_IF
	ELSE
		IF stValue.fValue <= i_fThreshold THEN
			iq_bCond := TRUE;
		ELSIF stValue.fValue > i_fThreshold + i_stSet.fHyst THEN
			iq_bCond := FALSE;
		END_IF
	END_IF
END_IF
M_Judge := iq_bCond;
END_METHOD

METHOD M_CheckSet : WSTRING(63)		// 설정 점검: 해소 폭 (FB_RuleBit은 점검할 값 없음)
M_CheckSet := "";
IF NOT F_RealOk(i_stSet.fHyst) THEN	// [결함 13 수정 2026-11-04]
	M_CheckSet := "해소 폭 fHyst 숫자 아님";
ELSIF i_stSet.fHyst < 0.0 THEN
	M_CheckSet := "해소 폭 fHyst 음수";
END_IF
END_METHOD

END_FUNCTION_BLOCK

// ---- 20_Module/Common/FB_BreakerCtrl.TcPOU
FUNCTION_BLOCK FB_BreakerCtrl EXTENDS FB_ModuleBase IMPLEMENTS I_OutputRule, I_ProtectionRule	// 차단기(VCB) 운전원 투입·개방: 지령 → 코일 펄스(DO) → 상태 접점 확인 → 실패 감시
// 출력: 출력 규칙 칸 두 개에 같은 인스턴스를 등록하고 g_astOutputCfg의 fThreshold로 코일을 고름 (1 = 투입 코일, 2 = 개방 코일). 장비·점은 그 칸의 nAux·nPoint, 지연 0·유지 끔
// 실패 감시: 보호 규칙 칸에도 같은 인스턴스를 등록 (g_astRuleCfg 조치 None이면 알람만). 조건 = 투입 실패 또는 개방 실패 (다음 성공 조작 또는 i_bResetFail로 풀림)
// 지령: HMI가 i_bCloseCmd·i_bOpenCmd를 켬 (상승 에지 1번에 1회). 같이 오면 개방이 이김. 투입은 상태 접점이 정상이고 개방 상태일 때만, 개방은 언제나 (조작 중이어도 끼어듦)
// 보호 트립 같은 자동 개방은 다른 출력 규칙(FB_RuleBit 등)을 같은 개방 코일 점에 등록 (같은 점은 OR)
// 스캔마다 한 번만 갱신 (보호 규칙·출력 규칙으로 여러 번 불려도 첫 호출에서만)
VAR_INPUT
	i_ipAux			: I_AuxDevice;		// 상태 접점을 읽을 보조 장비 (선언 때 지정)
	i_nClosedPoint	: UINT;				// 디지털 입력 점: TRUE = 투입 상태
	i_stSet			: ST_BreakerSet;	// 펄스 폭·확인 시간 (MAIN A_PassModuleSet이 g_stModuleSet 칸을 넘김. 안 넘기면 기본값)
	i_bCloseCmd		: BOOL;				// 투입 지령 (HMI, 상승 에지)
	i_bOpenCmd		: BOOL;				// 개방 지령 (HMI, 상승 에지)
	i_bResetFail	: BOOL;				// 실패 표시 풀기 (HMI, 상승 에지)
END_VAR
VAR_OUTPUT
	q_bClosed		: BOOL;		// 투입 상태 (상태 접점, 마지막으로 읽은 값)
	q_bStateValid	: BOOL;		// 상태 접점을 읽을 수 있음 (보조 장비 통신 정상)
	q_bClosePulse	: BOOL;		// 투입 코일 출력 중
	q_bOpenPulse	: BOOL;		// 개방 코일 출력 중
	q_bBusy			: BOOL;		// 조작 확인 중
	q_bCloseFail	: BOOL;		// 투입 실패 (확인 시간 안에 투입 상태가 안 됨)
	q_bOpenFail		: BOOL;		// 개방 실패
END_VAR
VAR
	_rtClose		: R_TRIG;
	_rtOpen			: R_TRIG;
	_rtReset		: R_TRIG;
	_tonPulse		: TON;
	_tonConfirm		: TON;
	_nOp			: INT;		// 진행 중인 조작 (OP_NONE / OP_CLOSE / OP_OPEN)
	_fbTask			: GETCURTASKINDEX;
	_nLastCycle		: UDINT;
	_bRan			: BOOL;
END_VAR
VAR CONSTANT
	OP_NONE			: INT := 0;
	OP_CLOSE		: INT := 1;
	OP_OPEN			: INT := 2;
	COIL_CLOSE		: REAL := 1.0;	// 출력 규칙 fThreshold: 투입 코일
	COIL_OPEN		: REAL := 2.0;	// 개방 코일
	RSN_CLOSE_FAIL	: UINT := 1;
	RSN_OPEN_FAIL	: UINT := 2;
END_VAR

METHOD PRIVATE M_Update		// 스캔마다 한 번: 상태 읽기 → 지령 → 펄스 → 확인
VAR
	nCycle	: UDINT;
	bNew	: BOOL;
END_VAR
_fbTask();
nCycle := TwinCAT_SystemInfoVarList._TaskInfo[_fbTask.index].CycleCount;
IF _bRan AND nCycle = _nLastCycle THEN
	RETURN;		// 이번 스캔은 이미 갱신함
END_IF
_bRan		:= TRUE;
_nLastCycle	:= nCycle;

// 상태 접점
q_bStateValid := FALSE;
IF i_ipAux <> 0 THEN
	q_bStateValid := i_ipAux.Comm;
	IF q_bStateValid THEN
		q_bClosed := i_ipAux.M_GetBit(i_nClosedPoint);
	END_IF
END_IF

// 지령 (개방이 이김. 투입은 상태를 알고 개방 상태일 때만, 진행 중인 조작이 없을 때만)
_rtClose(CLK := i_bCloseCmd);
_rtOpen(CLK := i_bOpenCmd);
_rtReset(CLK := i_bResetFail);
IF _rtReset.Q THEN
	q_bCloseFail	:= FALSE;
	q_bOpenFail		:= FALSE;
END_IF
bNew := FALSE;
IF _rtOpen.Q AND NOT (q_bStateValid AND NOT q_bClosed) THEN
	_nOp	:= OP_OPEN;
	bNew	:= TRUE;
ELSIF _rtClose.Q AND _nOp = OP_NONE AND q_bStateValid AND NOT q_bClosed THEN
	_nOp	:= OP_CLOSE;
	bNew	:= TRUE;
END_IF
IF bNew THEN
	_tonPulse(IN := FALSE);
	_tonConfirm(IN := FALSE);
END_IF

// 펄스·확인
_tonPulse(IN := _nOp <> OP_NONE, PT := i_stSet.tPulse);
_tonConfirm(IN := _nOp <> OP_NONE, PT := i_stSet.tConfirm);
q_bClosePulse	:= _nOp = OP_CLOSE AND NOT _tonPulse.Q;
q_bOpenPulse	:= _nOp = OP_OPEN AND NOT _tonPulse.Q;
IF _nOp = OP_CLOSE THEN
	IF q_bStateValid AND q_bClosed THEN
		_nOp			:= OP_NONE;
		q_bCloseFail	:= FALSE;
	ELSIF _tonConfirm.Q THEN
		_nOp			:= OP_NONE;
		q_bCloseFail	:= TRUE;
	END_IF
ELSIF _nOp = OP_OPEN THEN
	IF q_bStateValid AND NOT q_bClosed THEN
		_nOp			:= OP_NONE;
		q_bOpenFail		:= FALSE;
	ELSIF _tonConfirm.Q THEN
		_nOp			:= OP_NONE;
		q_bOpenFail		:= TRUE;
	END_IF
END_IF
q_bBusy := _nOp <> OP_NONE;
END_METHOD

METHOD M_Check : BOOL		// 출력 규칙: fThreshold 1 = 투입 코일, 2 = 개방 코일
VAR_INPUT
	i_fThreshold	: REAL;
END_VAR
M_Update();
IF i_fThreshold = COIL_CLOSE THEN
	M_Check := q_bClosePulse;
ELSIF i_fThreshold = COIL_OPEN THEN
	M_Check := q_bOpenPulse;
ELSE
	M_Check := FALSE;
END_IF
END_METHOD

METHOD M_Evaluate : BOOL		// 보호 규칙: 투입 실패 또는 개방 실패
VAR_INPUT
	i_stView	: ST_ProtView;	// 안 씀 (차단기 하나)
END_VAR
M_Update();
M_Evaluate := q_bCloseFail OR q_bOpenFail;
END_METHOD

METHOD M_ReasonText : WSTRING(63)
VAR_INPUT
	i_nReason	: UINT;
END_VAR
CASE i_nReason OF
	RSN_CLOSE_FAIL:	M_ReasonText := "차단기 투입 실패";
	RSN_OPEN_FAIL:	M_ReasonText := "차단기 개방 실패";
ELSE
	M_ReasonText := WCONCAT("이유 ", TO_WSTRING(i_nReason));
END_CASE
END_METHOD

METHOD M_CheckSet : WSTRING(63)		// 설정 점검: 펄스 폭, 확인 시간
M_CheckSet := "";
IF i_stSet.tPulse = T#0S THEN
	M_CheckSet := "펄스 폭 tPulse 0";
ELSIF i_stSet.tConfirm < i_stSet.tPulse THEN
	M_CheckSet := "확인 시간 tConfirm이 펄스 폭보다 짧음";
END_IF
END_METHOD

END_FUNCTION_BLOCK

// ---- 20_Module/Virtual/FB_BmsSim.TcPOU
FUNCTION_BLOCK FB_BmsSim EXTENDS FB_DeviceBase IMPLEMENTS I_Bms		// 가상 배터리 (시험용)
VAR_INPUT
	i_fPDc			: REAL;				// kW, 배터리에서 나가는 전력 (방전 +). PRG_SimLink가 넣음
	i_fSocInit		: REAL := 50.0;		// %
	i_fCapacity		: REAL := 4000.0;	// kWh
	i_fPLimit		: REAL := 2000.0;	// kW, 충·방전 한도
	i_bForceFault	: BOOL;				// 시험: 배터리 고장
	i_bForceSysStop	: BOOL;				// 시험: 시스템 정지
	i_bForceCommLoss	: BOOL;			// 시험: 응답 안 함. i_tCommTimeout 뒤 통신 이상
	i_bIgnoreCmd	: BOOL;				// 시험: 상태 명령을 접수하되 접촉기는 바꾸지 않음
	i_bDisableAutoOpen : BOOL;		// 시험: 고장·시스템 정지 때 자동 개방 안 함 (명령에 의한 개방은 별도)
END_VAR
VAR
	_bInit			: BOOL;
	_bClosed		: BOOL;
	_fSoc			: REAL;
	_stBat			: ST_BatState;
END_VAR

PROPERTY BatState : ST_BatState
GET
BatState := _stBat;
END_GET
END_PROPERTY

METHOD M_Cycle
VAR
	fDtHour		: REAL;
END_VAR
IF M_IsReadTime() AND NOT i_bForceCommLoss THEN		// 시험: 통신 끊김이면 응답 안 함
	M_MarkAlive();
END_IF
M_UpdateComm();

IF NOT _bInit THEN
	_fSoc	:= i_fSocInit;
	_bInit	:= TRUE;
END_IF

// 고장·시스템 정지면 접촉기 개방 (시험 입력으로 자동 개방만 끌 수 있음)
IF (i_bForceFault OR i_bForceSysStop) AND NOT i_bDisableAutoOpen THEN
	_bClosed := FALSE;
END_IF

// SOC 적분 (접촉기 투입 중일 때만)
IF _bClosed AND i_fCapacity > 0 THEN
	fDtHour	:= F_CycleSec() / 3600.0;
	_fSoc	:= LIMIT(0.0, _fSoc - i_fPDc * fDtHour / i_fCapacity * 100.0, 100.0);
END_IF

_stBat.bComm			:= _bComm;
_stBat.bContactorClosed	:= _bClosed;
_stBat.bWarn			:= FALSE;
_stBat.bFault			:= i_bForceFault;
_stBat.bSysStop			:= i_bForceSysStop;
_stBat.stSoc.fValue		:= _fSoc;
_stBat.stSoc.bValid		:= TRUE;
_stBat.stSoh.fValue		:= 100.0;
_stBat.stSoh.bValid		:= TRUE;
_stBat.fPChgMax			:= SEL(_fSoc < 100.0, 0.0, i_fPLimit);
_stBat.fPDisMax			:= SEL(_fSoc > 0.0, 0.0, i_fPLimit);
END_METHOD

METHOD M_SetStateCmd : BOOL
VAR_INPUT
	i_stCmd		: ST_BatCmd;
END_VAR
CASE i_stCmd.eCmd OF
	E_BatCmd.Close:
		IF NOT i_bIgnoreCmd AND NOT i_bForceFault AND NOT i_bForceSysStop THEN _bClosed := TRUE; END_IF
	E_BatCmd.Open,
	E_BatCmd.EStop:
		IF NOT i_bIgnoreCmd THEN _bClosed := FALSE; END_IF
	E_BatCmd.Reset:
		;	// 가상 장비는 고장 리셋을 입력(i_bForceFault)으로 함
ELSE
	RETURN;
END_CASE
M_SetStateCmd := TRUE;
END_METHOD

END_FUNCTION_BLOCK

// ---- 20_Module/Ups/FB_UpsChargeRequest.TcPOU
FUNCTION_BLOCK FB_UpsChargeRequest // 요청 번호와 완료 확인 관리
VAR_INPUT
 i_eAction : E_UpsChargeAction;
 i_fValue : REAL;
 i_tTimeout : TIME;
 i_stFeedback : ST_UpsChargeFeedback;
END_VAR
VAR_OUTPUT
 q_stRequest : ST_UpsChargeRequest;
 q_bDone : BOOL;
 q_bError : BOOL;
END_VAR
VAR
 _nSeq : UDINT;
 _ton : TON;
 _bWasPending : BOOL;
END_VAR

_bWasPending := q_stRequest.bValid;
IF i_eAction = E_UpsChargeAction.NoRequest THEN
 q_stRequest.bValid := FALSE;
 q_bDone := FALSE;
 q_bError := FALSE;
ELSE
 IF NOT q_stRequest.bValid AND NOT q_bDone AND NOT q_bError THEN
  _nSeq := F_UpsNextSeq(_nSeq);
  q_stRequest.nSeq := _nSeq;
  q_stRequest.eAction := i_eAction;
  q_stRequest.fValue := i_fValue;
  q_stRequest.bValid := TRUE;
 END_IF
 IF _bWasPending AND i_stFeedback.bValid AND i_stFeedback.nSeq = q_stRequest.nSeq THEN
  q_stRequest.bValid := FALSE;
  q_bDone := i_stFeedback.bConfirmed;
  q_bError := NOT i_stFeedback.bConfirmed;
 END_IF
END_IF
_ton(IN:=q_stRequest.bValid, PT:=i_tTimeout);
IF q_stRequest.bValid AND (_ton.Q OR i_tTimeout = T#0MS) THEN
 q_stRequest.bValid := FALSE;
 q_bError := TRUE;
END_IF

END_FUNCTION_BLOCK

// ---- 20_Module/Ups/FB_UpsChargeSequence.TcPOU
FUNCTION_BLOCK FB_UpsChargeSequence // 충방전 순서에 따른 요청 생성
VAR_INPUT
 i_bEnable : BOOL;
 i_bCancel : BOOL;
 i_bReset : BOOL;
 i_bResetReference : BOOL; // 기준 결과 초기화
 i_eMode : E_UpsChargeMode;
 i_stSet : ST_UpsChargeSet;
 i_stUps : ST_UpsState;
 i_stBms : ST_EsolutionState;
 i_stTime : ST_LocalTime;
 i_stFeedback : ST_UpsChargeFeedback;
END_VAR
VAR_OUTPUT
 q_eStep : E_UpsChargeStep;
 q_eMode : E_UpsChargeMode;
 q_stRequest : ST_UpsChargeRequest;
 q_stActiveSet : ST_UpsChargeSet; // 이번 운전에 고정한 설정
 q_bDone : BOOL; // 정상 완료
 q_bCanceled : BOOL; // 취소 완료
 q_bConflict : BOOL; // 다른 주 운전 시작 충돌
 q_bRecoveryRequired : BOOL; // 현장 상태 확인 필요
 q_nError : UINT; // 1: 설정, 2: 통신/보호, 3: 요청, 4: 모드, 5: 시간 초과
 q_bReferenceValid : BOOL; // 최초 주기적 방전 결과
 q_fReferenceStartVoltageV : REAL;
 q_fReferenceEndVoltageV : REAL;
 q_stReferenceTime : ST_LocalTime;
 q_fStartVoltageV : REAL;
 q_fEndVoltageV : REAL;
 q_stLastTime : ST_LocalTime;
 q_nLastScheduleDate : UDINT;
END_VAR
VAR
 _fbRequest : FB_UpsChargeRequest;
 _eAction : E_UpsChargeAction;
 _bNormal : BOOL;
 _bDataOk : BOOL;
 _bStarted : BOOL;
 _bCanceled : BOOL;
 _bClearRequest : BOOL;
 _bUpsDischargeRequested : BOOL;
 _bDue : BOOL;
 _bEndReached : BOOL;
 _bRestartReached : BOOL;
 _nDate : UDINT;
 _nWeek : UINT;
 _nModeSample : UDINT;
 _tonExtra : TON;
 _tonRest : TON;
 _tonInitial : TON;
 _tonDischarge : TON;
 _tonRun : TON;
 _tonMode : TON;
 _tonAbnormal : TON; // 운전 중 BBC Normal 해제가 이어진 시간
 _bProtTrip : BOOL; // 사고/고장 3~6단계 신호 (동작시퀀스 7쪽)
 _bHardOk : BOOL; // 데이터 유효, 3~6단계·BMS Minor 없음
 _bActive : BOOL; // 운전 단계 (Idle·WaitNormal·Complete·Fault 아님)
 _bWaitStep : BOOL; // 오래 기다리는 단계 (스케줄 대기·휴지)
 _bSafeCancel : BOOL; // 고장 뒤 UPS 방전 취소 요청 중
 _nNewFault : UINT; // 이번 스캔에 생긴 고장 번호
END_VAR

q_bDone := FALSE;
q_bCanceled := FALSE;
IF i_bResetReference AND (q_eStep = E_UpsChargeStep.Idle OR q_eStep = E_UpsChargeStep.WaitSchedule) THEN
 q_bReferenceValid:=FALSE;
END_IF
_eAction := E_UpsChargeAction.NoRequest;
_bClearRequest := FALSE;
_nNewFault := 0;
_bDataOk := i_stUps.bValid AND i_stBms.bValid;
// 동작시퀀스 7쪽 3~6단계: UPS·BMS가 배터리 컨버터 정지·MCCB Trip·컨택터 차단을 하는 상황. 어느 단계에서든 즉시 고장, 자동 재개 없음
// 비상정지(6), BMS Major(3), STATUS2 b12·b13 RCD 1·2단계 = DC전로 지락(3·4), b14 화재(5), BBC 정지 알람(4), BMS 고장·잠금(5)
_bProtTrip := (i_stUps.bValid AND (i_stUps.bEmergencyStop OR i_stUps.bBmsMajor
  OR (i_stUps.wStatus2 AND 16#7000) <> 0 OR (i_stUps.wBbcAlarm AND 16#0FA8) <> 0))
 OR (i_stBms.bValid AND (i_stBms.bFault OR i_stBms.bSystemLock));
// 2단계 BMS Minor(충전만 차단)와 통신 장애(15쪽: 정상운전 + 점검 요청)도 운전 단계는 멈추지만, 대기 단계에서는 기다림만
_bHardOk := _bDataOk AND NOT _bProtTrip AND NOT i_stUps.bBmsMinor;
// Rect Normal 0 = 정전·정류부 중고장(3단계) → 운전 단계 즉시 고장. BBC Normal은 BBC 기동 직후 3초 과도 구간에 0 → tModeTimeout 넘게 이어질 때만 고장
_bNormal := _bHardOk AND i_stUps.bRectNormal AND i_stUps.bBbcNormal;
_bActive := q_eStep <> E_UpsChargeStep.Idle AND q_eStep <> E_UpsChargeStep.WaitNormal
 AND q_eStep <> E_UpsChargeStep.Complete AND q_eStep <> E_UpsChargeStep.Fault;
// 스케줄 대기(최대 한 달)·휴지(30일)는 3~6단계만 고장. 그 밖의 이상은 고장으로 보지 않고 다음 단계로 넘어가지 않음
_bWaitStep := q_eStep = E_UpsChargeStep.WaitSchedule OR q_eStep = E_UpsChargeStep.Rest;
_tonAbnormal(IN:=_bActive AND NOT _bWaitStep AND _bHardOk AND i_stUps.bRectNormal AND NOT i_stUps.bBbcNormal,
 PT:=q_stActiveSet.tModeTimeout);
q_bConflict := q_eMode <> E_UpsChargeMode.Off AND i_eMode <> q_eMode AND i_eMode <> E_UpsChargeMode.Off;
IF i_bReset AND NOT i_bEnable AND (q_eStep = E_UpsChargeStep.Fault OR q_eStep = E_UpsChargeStep.Complete) THEN
 // 리셋은 현장 확인 후 수행. 장비를 정지시키는 명령이 아님.
 q_eStep := E_UpsChargeStep.Idle;
 q_eMode := E_UpsChargeMode.Off;
 q_nError := 0;
 q_bRecoveryRequired := FALSE;
 _bStarted := FALSE;
 _bSafeCancel := FALSE;
END_IF

IF _bActive THEN
 IF _bProtTrip OR (NOT _bWaitStep AND (NOT _bHardOk OR NOT i_stUps.bRectNormal OR _tonAbnormal.Q)) THEN
  _nNewFault := 2;
 ELSIF _fbRequest.q_bError THEN
  _nNewFault := 3;
 ELSIF NOT i_bEnable OR i_bCancel OR i_eMode = E_UpsChargeMode.Off THEN
  IF NOT _bCanceled THEN
   _bCanceled := TRUE;
   _bClearRequest := TRUE;
   IF NOT _bStarted THEN
    q_eStep := E_UpsChargeStep.Complete;
   ELSIF q_eMode = E_UpsChargeMode.Trickle THEN
    q_eStep := E_UpsChargeStep.BbcResume;
   ELSIF _bUpsDischargeRequested THEN
    q_eStep := E_UpsChargeStep.CancelUps;
   ELSE
    q_eStep := E_UpsChargeStep.CancelBms;
   END_IF
  END_IF
 END_IF
END_IF

_bEndReached := i_stUps.fBatteryVoltageV >= q_stActiveSet.fEndVoltageV;
_bRestartReached := i_stUps.fBatteryVoltageV <= q_stActiveSet.fStartVoltageV;
IF q_stActiveSet.nTrickleCriterion = 2 THEN
 _bEndReached := i_stBms.fSocPct >= q_stActiveSet.fEndSocPct;
 _bRestartReached := i_stBms.fSocPct <= q_stActiveSet.fStartSocPct;
END_IF
_tonExtra(IN:=q_eStep = E_UpsChargeStep.ExtraCharge, PT:=q_stActiveSet.tExtraCharge);
_tonRest(IN:=q_eStep = E_UpsChargeStep.Rest, PT:=q_stActiveSet.tRestart);
_tonInitial(IN:=q_eStep = E_UpsChargeStep.ExtraCharge AND q_eMode = E_UpsChargeMode.Periodic, PT:=q_stActiveSet.tInitialCharge);
_tonDischarge(IN:=q_eStep = E_UpsChargeStep.Running AND q_eMode = E_UpsChargeMode.Periodic, PT:=q_stActiveSet.tPeriodicDischarge);
_tonRun(IN:=q_eStep = E_UpsChargeStep.Running, PT:=q_stActiveSet.tRunTimeout);
_tonMode(IN:=q_eStep = E_UpsChargeStep.WaitRunning OR q_eStep = E_UpsChargeStep.WaitReady
 OR q_eStep = E_UpsChargeStep.WaitFloat, PT:=q_stActiveSet.tModeTimeout);
IF _nNewFault = 0 AND _tonMode.Q THEN _nNewFault:=4; END_IF
IF _nNewFault = 0 AND _tonRun.Q THEN _nNewFault:=5; END_IF
IF _nNewFault <> 0 THEN
 // UPS 방전을 요청하고 끝내지 못한 채 고장이면 방전 취소를 한 번 요청 (주기적 방전은 취소 전까지 계속됨)
 _bSafeCancel := _bUpsDischargeRequested AND (q_eStep = E_UpsChargeStep.StartDischarge
  OR q_eStep = E_UpsChargeStep.WaitRunning OR q_eStep = E_UpsChargeStep.Running OR q_eStep = E_UpsChargeStep.CancelUps);
 q_nError := _nNewFault;
 q_bRecoveryRequired := _bStarted OR _nNewFault = 5;
 _bClearRequest := TRUE; // 이전 요청의 확인·오류를 취소 요청에 다시 쓰지 않음
 q_eStep := E_UpsChargeStep.Fault;
END_IF

_bDue := FALSE;
IF i_stTime.bValid AND i_stTime.nMonth >= 1 AND i_stTime.nMonth <= 12
 AND i_stTime.nDay >= 1 AND i_stTime.nDay <= 31 THEN
 _nDate := UINT_TO_UDINT(i_stTime.nYear)*10000 + UINT_TO_UDINT(i_stTime.nMonth)*100 + UINT_TO_UDINT(i_stTime.nDay);
 _nWeek := (i_stTime.nDay-1)/7+1;
 _bDue := (q_stActiveSet.wMonthMask AND SHL(WORD#1,i_stTime.nMonth-1)) <> 0
  AND _nWeek = q_stActiveSet.nWeek AND i_stTime.nDayOfWeek = q_stActiveSet.nWeekDay
  AND i_stTime.nHour = q_stActiveSet.nHour AND _nDate > q_nLastScheduleDate;
END_IF

IF NOT _bClearRequest THEN
CASE q_eStep OF
 E_UpsChargeStep.Idle:
  IF i_bEnable AND NOT i_bCancel AND NOT i_bReset AND i_eMode <> E_UpsChargeMode.Off THEN
   q_eMode:=i_eMode; q_stActiveSet:=i_stSet; q_nError:=0;
   _bCanceled:=FALSE; _bStarted:=FALSE; _bUpsDischargeRequested:=FALSE;
   q_eStep:=E_UpsChargeStep.WaitNormal;
  END_IF
 E_UpsChargeStep.WaitNormal:
  IF NOT i_bEnable OR i_bCancel OR i_eMode = E_UpsChargeMode.Off THEN
   _bCanceled:=TRUE; q_eStep:=E_UpsChargeStep.Complete;
  ELSIF _bNormal THEN
   IF i_stUps.nBatMode <> 0 THEN
    q_bConflict:=TRUE;
   ELSIF q_stActiveSet.tRequestTimeout = T#0MS OR q_stActiveSet.tModeTimeout = T#0MS THEN
    q_nError:=1; q_eStep:=E_UpsChargeStep.Fault;
   ELSE
    CASE q_eMode OF
     E_UpsChargeMode.Trickle:
      IF (q_stActiveSet.nTrickleCriterion = 1 AND q_stActiveSet.fStartVoltageV > 0.0
       AND q_stActiveSet.fEndVoltageV > q_stActiveSet.fStartVoltageV)
       OR (q_stActiveSet.nTrickleCriterion = 2 AND q_stActiveSet.fStartSocPct >= 0.0
       AND q_stActiveSet.fEndSocPct > q_stActiveSet.fStartSocPct AND q_stActiveSet.fEndSocPct <= 100.0) THEN
       IF q_stActiveSet.tExtraCharge > T#0MS AND q_stActiveSet.tRestart > T#0MS THEN
        q_eStep:=E_UpsChargeStep.BbcStart;
       ELSE q_nError:=1; q_eStep:=E_UpsChargeStep.Fault; END_IF
      ELSE q_nError:=1; q_eStep:=E_UpsChargeStep.Fault; END_IF
     E_UpsChargeMode.Periodic:
      IF q_stActiveSet.fFloatVoltageV > 0.0 AND q_stActiveSet.fPeriodicCurrentA > 0.0
       AND q_stActiveSet.tInitialCharge > T#0MS AND q_stActiveSet.tPeriodicDischarge > T#0MS AND q_stActiveSet.tRunTimeout > q_stActiveSet.tPeriodicDischarge
       AND q_stActiveSet.wMonthMask <> 0 AND q_stActiveSet.wMonthMask <= 16#0FFF
       AND q_stActiveSet.nWeek >= 1 AND q_stActiveSet.nWeek <= 4
       AND q_stActiveSet.nWeekDay <= 6 AND q_stActiveSet.nHour <= 23 THEN
       q_eStep:=E_UpsChargeStep.WaitSchedule;
      ELSE q_nError:=1; q_eStep:=E_UpsChargeStep.Fault; END_IF
     E_UpsChargeMode.Pulse:
      IF q_stActiveSet.fPulseChargeA > 0.0 AND q_stActiveSet.fPulseDischargeA > 0.0
       AND q_stActiveSet.tPulseCharge > T#0MS AND q_stActiveSet.tPulseDischarge > T#0MS
       AND q_stActiveSet.nPulseCycles > 0 AND q_stActiveSet.tRunTimeout > T#0MS
       AND (UDINT_TO_LREAL(TIME_TO_UDINT(q_stActiveSet.tPulseCharge))
       + UDINT_TO_LREAL(TIME_TO_UDINT(q_stActiveSet.tPulseDischarge)))
       *UINT_TO_LREAL(q_stActiveSet.nPulseCycles) < UDINT_TO_LREAL(TIME_TO_UDINT(q_stActiveSet.tRunTimeout)) THEN
       q_eStep:=E_UpsChargeStep.PrepareBms;
      ELSE q_nError:=1; q_eStep:=E_UpsChargeStep.Fault; END_IF
     ELSE q_nError:=1; q_eStep:=E_UpsChargeStep.Fault;
    END_CASE
   END_IF
  END_IF
 E_UpsChargeStep.WaitSchedule:
  IF _bDue AND i_stUps.nBatMode = 0 AND _bNormal THEN
   q_nLastScheduleDate:=_nDate;
   IF i_stUps.fBatteryVoltageV <= q_stActiveSet.fFloatVoltageV THEN q_eStep:=E_UpsChargeStep.ExtraCharge;
   ELSE q_eStep:=E_UpsChargeStep.PrepareBms; END_IF
  END_IF
 E_UpsChargeStep.BbcStart:
  IF _fbRequest.q_bDone THEN q_eStep:=E_UpsChargeStep.WaitEnd;
  ELSE _eAction:=E_UpsChargeAction.BbcOn; _bStarted:=TRUE; END_IF
 E_UpsChargeStep.WaitEnd:
  IF _bEndReached THEN q_eStep:=E_UpsChargeStep.ExtraCharge; END_IF
 E_UpsChargeStep.ExtraCharge:
  IF q_eMode = E_UpsChargeMode.Trickle AND _tonExtra.Q THEN q_eStep:=E_UpsChargeStep.BbcReady;
  ELSIF q_eMode = E_UpsChargeMode.Periodic AND _tonInitial.Q THEN q_eStep:=E_UpsChargeStep.PrepareBms; END_IF
 E_UpsChargeStep.BbcReady:
  IF _fbRequest.q_bDone THEN _nModeSample:=i_stUps.nSampleSeq; q_eStep:=E_UpsChargeStep.WaitReady;
  ELSE _eAction:=E_UpsChargeAction.BbcReady; END_IF
 E_UpsChargeStep.WaitReady:
  IF i_stUps.nSampleSeq <> _nModeSample AND i_stUps.nBatMode = 2 THEN q_eStep:=E_UpsChargeStep.Rest; END_IF
 E_UpsChargeStep.Rest:
  IF (_bRestartReached OR _tonRest.Q) AND _bHardOk AND i_stUps.bRectNormal THEN q_eStep:=E_UpsChargeStep.BbcStart; END_IF // 대기모드에서는 BBC Normal을 보지 않음
 E_UpsChargeStep.PrepareBms:
  IF i_stUps.nBatMode <> 0 THEN q_bConflict:=TRUE;
  ELSIF _fbRequest.q_bDone THEN q_eStep:=E_UpsChargeStep.StartDischarge;
  ELSE
   _bStarted:=TRUE;
   IF q_eMode = E_UpsChargeMode.Periodic THEN _eAction:=E_UpsChargeAction.BmsPreparePeriodic;
   ELSE _eAction:=E_UpsChargeAction.BmsPreparePulse; END_IF
  END_IF
 E_UpsChargeStep.StartDischarge:
  IF NOT _bUpsDischargeRequested AND i_stUps.nBatMode <> 0 THEN q_bConflict:=TRUE;
  ELSIF _fbRequest.q_bDone THEN _nModeSample:=i_stUps.nSampleSeq; q_eStep:=E_UpsChargeStep.WaitRunning;
  ELSE
   _bUpsDischargeRequested:=TRUE;
   IF q_eMode = E_UpsChargeMode.Periodic THEN _eAction:=E_UpsChargeAction.PeriodicStart;
   ELSE _eAction:=E_UpsChargeAction.PulseStart; END_IF
  END_IF
 E_UpsChargeStep.WaitRunning:
  IF i_stUps.nSampleSeq <> _nModeSample AND ((q_eMode = E_UpsChargeMode.Periodic AND i_stUps.nBatMode = 3)
   OR (q_eMode = E_UpsChargeMode.Pulse AND i_stUps.nBatMode = 4)) THEN
   q_fStartVoltageV:=i_stUps.fBatteryVoltageV;
   _nModeSample:=i_stUps.nSampleSeq; q_eStep:=E_UpsChargeStep.Running;
  END_IF
 E_UpsChargeStep.Running:
  IF (q_eMode = E_UpsChargeMode.Periodic AND i_stUps.nBatMode = 3) OR (q_eMode = E_UpsChargeMode.Pulse AND i_stUps.nBatMode = 4) THEN
   q_fEndVoltageV:=i_stUps.fBatteryVoltageV; // 방전 중 마지막 전압 = 종료 전압 (부동충전 복귀 뒤에는 전압이 다시 오름)
  END_IF
  IF i_stUps.nSampleSeq <> _nModeSample AND i_stUps.nBatMode = 0 THEN q_eStep:=E_UpsChargeStep.CancelBms;
  ELSIF q_eMode = E_UpsChargeMode.Periodic AND _tonDischarge.Q THEN q_eStep:=E_UpsChargeStep.CancelUps; END_IF
 E_UpsChargeStep.CancelUps:
  IF _fbRequest.q_bDone THEN q_eStep:=E_UpsChargeStep.CancelBms;
  ELSE _eAction:=E_UpsChargeAction.DischargeCancel; END_IF
 E_UpsChargeStep.CancelBms:
  IF _fbRequest.q_bDone THEN q_eStep:=E_UpsChargeStep.FloatRequest;
  ELSE _eAction:=E_UpsChargeAction.BmsDischargeCancel; END_IF
 E_UpsChargeStep.BbcResume:
  IF _fbRequest.q_bDone THEN q_eStep:=E_UpsChargeStep.FloatRequest;
  ELSE _eAction:=E_UpsChargeAction.BbcOn; END_IF
 E_UpsChargeStep.FloatRequest:
  IF _fbRequest.q_bDone THEN _nModeSample:=i_stUps.nSampleSeq; q_eStep:=E_UpsChargeStep.WaitFloat;
  ELSE _eAction:=E_UpsChargeAction.FloatCharge; END_IF
 E_UpsChargeStep.WaitFloat:
  IF i_stUps.nSampleSeq <> _nModeSample AND i_stUps.nBatMode = 0 THEN
   IF q_eMode = E_UpsChargeMode.Trickle THEN q_fEndVoltageV:=i_stUps.fBatteryVoltageV; END_IF
   q_stLastTime:=i_stTime; _bStarted:=FALSE; _bUpsDischargeRequested:=FALSE;
   IF _bCanceled THEN q_eStep:=E_UpsChargeStep.Complete;
   ELSIF q_eMode = E_UpsChargeMode.Periodic THEN
    IF NOT q_bReferenceValid THEN
     q_fReferenceStartVoltageV:=q_fStartVoltageV;
     q_fReferenceEndVoltageV:=q_fEndVoltageV;
     q_stReferenceTime:=i_stTime; q_bReferenceValid:=TRUE;
    END_IF
    q_bDone:=TRUE; q_eStep:=E_UpsChargeStep.WaitSchedule;
   ELSE q_bDone:=TRUE; q_eStep:=E_UpsChargeStep.Complete; END_IF
  END_IF
 E_UpsChargeStep.Complete:
  q_bCanceled:=_bCanceled;
  IF NOT i_bEnable THEN q_eStep:=E_UpsChargeStep.Idle; q_eMode:=E_UpsChargeMode.Off; END_IF
 E_UpsChargeStep.Fault:
  // 장비 보호·비상정지는 별도 담당. 자동 재시작하지 않음. 방전 중이었으면 UPS 데이터가 유효할 때 취소를 한 번 요청
  IF _bSafeCancel THEN
   IF _fbRequest.q_bDone OR _fbRequest.q_bError THEN _bSafeCancel:=FALSE;
   ELSIF i_stUps.bValid THEN _eAction:=E_UpsChargeAction.DischargeCancel; END_IF
  END_IF
END_CASE
END_IF
_fbRequest(i_eAction:=_eAction, i_fValue:=0.0, i_tTimeout:=q_stActiveSet.tRequestTimeout, i_stFeedback:=i_stFeedback);
q_stRequest:=_fbRequest.q_stRequest;

END_FUNCTION_BLOCK

// ---- 20_Module/Ups/FB_UpsTemperatureCharge.TcPOU
FUNCTION_BLOCK FB_UpsTemperatureCharge // 온도보상 전압 계산 및 적용 요청
VAR_INPUT
 i_bEnable : BOOL;
 i_bSuspend : BOOL;
 i_bReset : BOOL;
 i_stUps : ST_UpsState;
 i_stSet : ST_UpsChargeSet;
 i_stTime : ST_LocalTime;
 i_stFeedback : ST_UpsChargeFeedback;
END_VAR
VAR_OUTPUT
 q_stRequest : ST_UpsChargeRequest;
 q_fTargetVoltageV : REAL;
 q_fAppliedVoltageV : REAL;
 q_bSuspended : BOOL;
 q_bApplied : BOOL;
 q_nError : UINT; // 1: 설정/온도, 2: 통신/보호, 3: 적용 확인
 q_stLastTime : ST_LocalTime;
END_VAR
VAR
 _fbRequest : FB_UpsChargeRequest;
 _eAction : E_UpsChargeAction;
 _tonUpdate : TON;
 _bUpdateDone : BOOL;
 _bRestore : BOOL;
 _bWasSuspended : BOOL;
 _fPendingV : REAL;
 _bPending : BOOL;
END_VAR

_eAction:=E_UpsChargeAction.NoRequest;
q_bSuspended:=i_bSuspend OR i_stUps.nBatMode = 3 OR i_stUps.nBatMode = 4;
_tonUpdate(IN:=q_bApplied AND NOT _bUpdateDone, PT:=i_stSet.tTempUpdate);
_bUpdateDone:=FALSE;
IF i_bReset THEN q_nError:=0; END_IF
IF q_nError = 2 THEN q_nError:=0; END_IF // 통신·보호 이상은 래치하지 않음: 매 스캔 다시 판정, 풀리면 이어서 (Disable이면 부동충전 전압 복귀)
IF _fbRequest.q_bError THEN q_nError:=3; END_IF

IF q_nError = 0 AND (i_bEnable OR q_bApplied OR _bPending) THEN
 IF NOT i_stUps.bValid OR NOT i_stUps.bRectNormal OR NOT i_stUps.bBbcNormal
  OR i_stUps.bEmergencyStop OR i_stUps.bBmsMinor OR i_stUps.bBmsMajor
  OR (i_stUps.wStatus2 AND 16#7000) <> 0 OR (i_stUps.wBbcAlarm AND 16#0FA8) <> 0 THEN // RCD 1·2단계·화재, BBC 정지 알람 (동작시퀀스 7쪽)
  q_nError:=2; _bPending:=FALSE;
 ELSIF NOT (i_stSet.fBaseCellVoltageV > 0.0 AND i_stSet.nSeriesCells > 0
  AND i_stSet.fMinChargeVoltageV > 0.0
  AND i_stSet.fMaxChargeVoltageV >= i_stSet.fMinChargeVoltageV
  AND i_stSet.fMaxChargeVoltageV <= 6553.5
  AND i_stSet.fFloatVoltageV >= i_stSet.fMinChargeVoltageV
  AND i_stSet.fFloatVoltageV <= i_stSet.fMaxChargeVoltageV
  AND i_stSet.fMinTemperatureC < i_stSet.fMaxTemperatureC
  AND i_stSet.tRequestTimeout > T#0MS AND i_stSet.tTempUpdate > T#0MS) THEN
  q_nError:=1;
 ELSIF NOT q_bSuspended THEN
  IF NOT _bPending THEN
   _bRestore:=NOT i_bEnable;
   IF _bRestore THEN q_fTargetVoltageV:=i_stSet.fFloatVoltageV;
   ELSE
    IF i_stUps.fBatteryRoomTemperatureC < i_stSet.fMinTemperatureC
     OR i_stUps.fBatteryRoomTemperatureC > i_stSet.fMaxTemperatureC THEN q_nError:=1;
    ELSE q_fTargetVoltageV:=(i_stSet.fBaseCellVoltageV + i_stSet.fSlopeMvPerC*0.001
     *(i_stUps.fBatteryRoomTemperatureC-25.0))*UINT_TO_REAL(i_stSet.nSeriesCells); END_IF
   END_IF
   IF NOT (q_fTargetVoltageV >= i_stSet.fMinChargeVoltageV AND q_fTargetVoltageV <= i_stSet.fMaxChargeVoltageV) THEN q_nError:=1; END_IF
   // 주기 갱신은 전압이 레지스터 해상도(0.1 V) 이상 바뀔 때만 씀. 아니면 쓰지 않고 주기만 다시 시작
   IF q_nError = 0 AND (NOT q_bApplied OR _bRestore OR _bWasSuspended
    OR (_tonUpdate.Q AND ABS(q_fTargetVoltageV - q_fAppliedVoltageV) >= 0.1)) THEN
    _fPendingV:=q_fTargetVoltageV; _bPending:=TRUE;
   ELSIF _tonUpdate.Q THEN
    _bUpdateDone:=TRUE;
   END_IF
  END_IF
  IF _bPending AND q_nError = 0 THEN
   IF _fbRequest.q_bDone THEN
    q_fAppliedVoltageV:=_fPendingV; q_stLastTime:=i_stTime;
    q_bApplied:=NOT _bRestore; _bPending:=FALSE; _bUpdateDone:=TRUE;
   ELSE _eAction:=E_UpsChargeAction.ChargeVoltage; END_IF
  END_IF
 END_IF
END_IF
IF q_bSuspended THEN _bPending:=FALSE; END_IF
_bWasSuspended:=q_bSuspended;
_fbRequest(i_eAction:=_eAction, i_fValue:=_fPendingV, i_tTimeout:=i_stSet.tRequestTimeout, i_stFeedback:=i_stFeedback);
q_stRequest:=_fbRequest.q_stRequest;

END_FUNCTION_BLOCK

// ---- 20_Module/Driver/Bender/FB_BenderIso685.TcPOU
FUNCTION_BLOCK FB_BenderIso685 EXTENDS FB_DeviceBase IMPLEMENTS I_AuxDevice		// Bender ISO685 절연감시장치(IMD) (Modbus TCP), 읽기 전용
(* ---------------------------------------------------------------
   기반: Helios FB_ISO685 v4.0. 동작만 옮기고 PmsStd 형식으로 다시 씀. 2026-11-09
   읽기: 읽기 주기마다 아래 묶음 하나씩 차례로 (Holding Register FC3, Helios와 같은 주소·수량)
     @MAP HR 4113  F32(앞 = 상위)  -  절연저항 측정값 (장치 단위, Helios도 배율 없음)
     @MAP HR 4115  U16  -  상위 바이트 = 시험 상태 (0 없음, 1 내부, 2 외부), 하위 바이트 = 알람 상태 (0 없음, 1 예비경고, 2 경고, 4 고장, 5 알람)
     @MAP HR 4273  F32  -  계통 연결 (system connection)
     @MAP HR 4289  F32  -  접지 연결 (connection to earth)
     @MAP HR 4305  F32  -  장치 오류 (device error)
     @MAP HR 4385  F32  -  대칭 절연 저하 (symmetric alarm)
     @MAP HR 12499 U32(앞 = 상위) ×2  -  응답값 1·2 (설정 경보값)
   점 (I_AuxDevice)
     AI 1 절연저항, 2 계통 연결, 3 접지 연결, 4 장치 오류, 5 대칭 절연 저하, 6 응답값 1, 7 응답값 2, 8 알람 상태 코드
     DI 1 경고 (알람 상태 2), DI 2 고장 (알람 상태 4), DI 3 시험 중
   Helios는 eIsoState로 "고장만" 또는 "경고 + 고장"을 보호 신호로 썼다 → PmsStd에서는 규칙(FB_RuleBit)에 DI 1·2 중 고를 점을 등록
   쓰기 없음. 맵 미확보: Helios 현장 기준, 펌웨어별 주소 확인 필요
   --------------------------------------------------------------- *)
VAR_INPUT
	i_bEnable		: BOOL;					// FALSE면 통신하지 않음 (장비 미설치)
	i_sIpAddr		: STRING(15);
	i_nPort			: UINT := 502;
	i_nUnitId		: BYTE := 1;
	i_tTimeout		: TIME := T#1S;
END_VAR
VAR
	_fbMbRead		: FB_MBReadRegs;
	_awBuf			: ARRAY[0..3] OF WORD;
	_bReadDue		: BOOL;					// 읽을 때가 됨 (매 스캔 M_IsReadTime)
	_bReading		: BOOL;
	_nBlock			: UINT;					// 지금 읽는 묶음 0..5
	_afAi			: ARRAY[1..8] OF REAL;
	_nAlarm			: WORD;					// 알람 상태 코드 (4115 하위 바이트)
	_nTest			: WORD;					// 시험 상태 (4115 상위 바이트)
	_bStatusOk		: BOOL;					// 묶음 0(측정값·상태)을 한 번이라도 읽음
END_VAR
VAR CONSTANT
	BLOCK_ADDR		: ARRAY[0..5] OF UINT := [4113, 4273, 4289, 4305, 4385, 12499];
	BLOCK_QTY		: ARRAY[0..5] OF UINT := [3, 2, 2, 2, 2, 4];
	ALARM_WARNING	: WORD := 2;
	ALARM_FAULT		: WORD := 4;
END_VAR

ACTION A_MapBlock:
CASE _nBlock OF
	0:
		_afAi[1]	:= F_WordsToReal(i_wHigh := _awBuf[0], i_wLow := _awBuf[1]);	// @MAP HR 4113 F32 절연저항
		_nAlarm		:= _awBuf[2] AND 16#00FF;										// @MAP HR 4115 하위 바이트 알람 상태
		_nTest		:= SHR(_awBuf[2], 8);											// @MAP HR 4115 상위 바이트 시험 상태
		_afAi[8]	:= WORD_TO_REAL(_nAlarm);
		_bStatusOk	:= TRUE;
	1:	_afAi[2]	:= F_WordsToReal(i_wHigh := _awBuf[0], i_wLow := _awBuf[1]);	// @MAP HR 4273 F32 계통 연결
	2:	_afAi[3]	:= F_WordsToReal(i_wHigh := _awBuf[0], i_wLow := _awBuf[1]);	// @MAP HR 4289 F32 접지 연결
	3:	_afAi[4]	:= F_WordsToReal(i_wHigh := _awBuf[0], i_wLow := _awBuf[1]);	// @MAP HR 4305 F32 장치 오류
	4:	_afAi[5]	:= F_WordsToReal(i_wHigh := _awBuf[0], i_wLow := _awBuf[1]);	// @MAP HR 4385 F32 대칭 절연 저하
	5:
		_afAi[6]	:= UDINT_TO_REAL(SHL(WORD_TO_UDINT(_awBuf[0]), 16) OR WORD_TO_UDINT(_awBuf[1]));	// @MAP HR 12499 U32 응답값 1
		_afAi[7]	:= UDINT_TO_REAL(SHL(WORD_TO_UDINT(_awBuf[2]), 16) OR WORD_TO_UDINT(_awBuf[3]));	// @MAP HR 12501 U32 응답값 2
END_CASE
END_ACTION

METHOD M_Cycle
_bReadDue := M_IsReadTime();
IF NOT _bReading THEN
	IF i_bEnable AND i_sIpAddr <> '' AND _bReadDue THEN
		_fbMbRead(sIPAddr := i_sIpAddr, nTCPPort := i_nPort, nUnitID := i_nUnitId,
			nQuantity := BLOCK_QTY[_nBlock], nMBAddr := BLOCK_ADDR[_nBlock], cbLength := BLOCK_QTY[_nBlock] * 2,
			pDestAddr := ADR(_awBuf), tTimeout := i_tTimeout, bExecute := TRUE);
		_bReading := TRUE;
	END_IF
ELSE
	_fbMbRead(bExecute := FALSE);
	IF NOT _fbMbRead.bBusy THEN
		IF NOT _fbMbRead.bError AND i_bEnable THEN
			A_MapBlock();
			M_MarkAlive();
		END_IF
		IF _nBlock >= 5 THEN _nBlock := 0; ELSE _nBlock := _nBlock + 1; END_IF
		_bReading := FALSE;
	END_IF
END_IF
M_UpdateComm();
END_METHOD

METHOD M_GetBit : BOOL		// DI 1 경고, 2 고장, 3 시험 중. 통신 이상이면 FALSE (규칙 FB_RuleBit은 Comm으로 따로 판단)
VAR_INPUT
	i_nPoint	: UINT;
END_VAR
IF Comm AND _bStatusOk THEN
	CASE i_nPoint OF
		1: M_GetBit := _nAlarm = ALARM_WARNING;
		2: M_GetBit := _nAlarm = ALARM_FAULT;
		3: M_GetBit := _nTest <> 0;
	END_CASE
END_IF
END_METHOD

METHOD M_GetValue : ST_Val		// AI 1..8 (머리 주석 참고)
VAR_INPUT
	i_nPoint	: UINT;
END_VAR
IF i_nPoint >= 1 AND i_nPoint <= 8 THEN
	M_GetValue.fValue := _afAi[i_nPoint];
	M_GetValue.bValid := Comm AND _bStatusOk;
END_IF
END_METHOD

METHOD M_SetBit		// 출력 없음
VAR_INPUT
	i_nPoint	: UINT;
	i_bValue	: BOOL;
END_VAR
;
END_METHOD

METHOD M_SetValue		// 출력 없음
VAR_INPUT
	i_nPoint	: UINT;
	i_fValue	: REAL;
END_VAR
;
END_METHOD

PROPERTY Comm : BOOL
GET
Comm := _bComm AND i_bEnable;
END_GET
END_PROPERTY

END_FUNCTION_BLOCK
